(* IEC 61131-3 sources: AutoPLC/data/rag_data/st/st_case_code (part 2) *)

(* ---- ELEMENT_GET.st ---- *)
FUNCTION ELEMENT_GET : string
VAR_INPUT
    SEP : BYTE;
    POS : INT;
END_VAR

VAR_IN_OUT
    ELEMENT : STRING[ELEMENT_LENGTH];
END_VAR_IN_OUT

VAR
    i : INT := 1;
    o : INT := 1;
    pt : POINTER TO ARRAY[1..ELEMENT_LENGTH] OF BYTE;
    po : POINTER TO ARRAY[1..ELEMENT_LENGTH] OF BYTE;
    cnt : INT;
    c : BYTE;
END_VAR
(* load pointers *)
pt := ADR(ELEMENT);
po := ADR(ELEMENT_GET);

(* search for the n-th occurence of a separation character and store position in i *)
WHILE (cnt < pos) AND (i < ELEMENT_LENGTH) AND (pt^[i] > 0) DO
	IF pt^[i] = sep THEN cnt := cnt + 1; END_IF;
	i := i + 1;
END_WHILE;

(* copy the list element to output *)
IF i < ELEMENT_LENGTH THEN c := pt^[i]; END_IF;
WHILE (c <> sep) AND (c > 0) AND (o < ELEMENT_LENGTH) AND (i < ELEMENT_LENGTH) DO
	po^[o] :=pt^[i];
	o := o + 1;
	i := i + 1;
	c := pt^[i];
END_WHILE;

(* terminate the output string *)
po^[o] := 0;

(* revision histroy
ks 05. apr. 2011	rev 1.0
	original release

*)
END_FUNCTION

(* ---- ELLIPSE_A.st ---- *)
FUNCTION ELLIPSE_A : REAL
VAR_INPUT
    R1: REAL;
    R2: REAL;
END_VAR
ELLIPSE_A := math.PI * R1 * R2;

(* revision histroy
hm	16. oct 2007	rev 1.0
	original version

hm	18. oct. 2008	rev 1.1
	using math constants
*)
END_FUNCTION

(* ---- ELLIPSE_C.st ---- *)
FUNCTION ELLIPSE_C : REAL
VAR_INPUT
    R1 : REAL;
    R2 : REAL;
END_VAR
ELLIPSE_C := math.PI * (3.0 * (R1+R2) - SQRT((3.0 * r1 + R2) * (3.0 * r2 + r1)));

(* revision histroy
hm	16. oct 2007	rev 1.0
	original version

hm	18. oct. 2008	rev 1.1
	using math constants

hm	10. mar. 2009	rev 1.2
	changed syntax of real constants to 0.0

*)
END_FUNCTION

(* ---- ERF.st ---- *)
FUNCTION ERF : REAL
VAR_INPUT
    X : REAL;
END_VAR_INPUT

VAR
    x2 : REAL;
    ax2 : REAL;
END_VAR
x2 := X*X;
ax2 := 0.147 * x2 + 1.0;
ERF := SQRT(1.0 - EXP(-X2 * ((0.27323954473516 + aX2)/(ax2)))) * SGN(x);

(* revision history
hm	7. apr. 2008	rev 1.0
	original version

hm	30. jun. 2008	rev 1.1
	added type conversions to avoid warnings under codesys 3.0

hm	25. oct. 2008	rev 1.2
	new code using new algorithm

hm	10. mar. 2009	rev 1.3
	real constants updated to new systax using dot
*)
END_FUNCTION

(* ---- ERFC.st ---- *)
FUNCTION ERFC : REAL
VAR_INPUT
    X : REAL;
END_VAR
ERFC := 1.0 - ERF(X);

(* revision history
hm	7. apr. 2008	rev 1.0
	original version

hm	10. mar. 2009	rev 1.1
	real constants updated to new systax using dot

*)
END_FUNCTION

(* ---- EVEN.st ---- *)
FUNCTION EVEN : BOOL
VAR_INPUT
    in : DINT; // Input variable declaration
END_VAR
EVEN := NOT in.0;

(* revision history
hm	1. oct 2006	rev 1.0
	ORIGINAL VERSION

hm	01.12.2007	rev 1.1
	changed code for improved performance

hm	21. mar. 2008	rev 1.2
	changed type of input IN from INT to DINT
*)
END_FUNCTION

(* ---- EXEC.st ---- *)
FUNCTION EXEC : string
VAR_INPUT
    str : STRING[STRING_LENGTH];
END_VAR

VAR
    pos : INT;
    R1 : REAL;
    R2 : REAL;
    operator : STRING[10];
END_VAR
(* extract both numbers and operator *)
EXEC := UPPERCASE(TRIM(str));

pos := FINDB_NONUM(EXEC);
IF pos > 1 THEN R1 := STRING_TO_REAL(LEFT(EXEC,pos-1)); END_IF;
R2 := STRING_TO_REAL(RIGHT(EXEC,LEN(EXEC)-pos));
EXEC := LEFT(EXEC,pos);
pos := FINDB_NUM(EXEC);
operator := RIGHT(EXEC,LEN(EXEC) - pos);
IF operator = '' AND LEN(str) = 0 THEN
	EXEC := '';
	RETURN;
ELSIF operator = '' THEN
	EXEC := str;
	RETURN;
END_IF;
IF operator = '^' THEN
	EXEC := REAL_TO_STRING(EXPT(R1, R2));
ELSIF operator = 'SQRT' THEN
	EXEC := REAL_TO_STRING(SQRT(R2));
ELSIF operator = 'SIN' THEN
	EXEC := REAL_TO_STRING(SIN(r2));
ELSIF operator = 'COS' THEN
	EXEC := REAL_TO_STRING(COS(r2));
ELSIF operator = 'TAN' THEN
	EXEC := REAL_TO_STRING(TAN(R2));
ELSIF operator = '*' THEN
	EXEC := REAL_TO_STRING(R1 * R2);
ELSIF operator = '/' THEN
	IF R2 <> 0 THEN EXEC := REAL_TO_STRING(R1 / R2); ELSE EXEC := 'ERROR'; END_IF;
ELSIF operator = '+' THEN
	EXEC := REAL_TO_STRING(r1 + r2);
ELSIF operator = '-' THEN
	EXEC := REAL_TO_STRING(r1 - r2);
ELSE
	EXEC := 'ERROR';
END_IF;

IF EXEC = 'ERROR' THEN
	RETURN;
(* some systems deliver integer instead of real *)
ELSIF FIND(EXEC,'.') = 0 THEN
	EXEC := CONCAT(EXEC, '.0');
(* some systems deliver n. instead of n.0 ! *)
ELSIF RIGHT(EXEC,1) = '.' THEN
	EXEC := CONCAT(EXEC,'0');
END_IF;

(* revision history

hm 	6.feb 2007		rev 1.1
	cos has to be written in uppercase
	divide by 0 will return an error

hm	5. mar. 2008	rev 1.2
	add a 0 to the string if a '.' is at the end of the string

hm	20. mar. 2008	rev 1.3
	make sure the function always returns a real value in the form of x.y

hm	29. mar. 2008	rev 1.4
	changed STRING to STRING(STRING_LENGTH)
*)
END_FUNCTION

(* ---- EXP10.st ---- *)
FUNCTION EXP10 : REAL
VAR_INPUT
    X : REAL;
END_VAR
EXP10 := EXP(X * 2.30258509299405);

(* revision history
hm	2. dec 2007		rev 1.0
	original version

*)
END_FUNCTION

(* ---- EXPN.st ---- *)
FUNCTION EXPN : REAL
VAR_INPUT
    X : REAL;  // Input variable of type REAL
    N : INT;   // Input variable of type INT
END_VAR

VAR
    sign : BOOL;  // Local variable of type BOOL
END_VAR
sign := n.15;
N := ABS(N);
IF N.0 THEN EXPN := X; ELSE EXPN := 1.0; END_IF;
N := SHR(N,1);
WHILE N > 0 DO
   X := X * X;
   IF N.0 THEN EXPN := EXPN * X; END_IF;
   N := SHR(N,1);
END_WHILE;
IF sign THEN EXPN := 1.0 / EXPN; END_IF;

(* revision history
hm	4. dec 2007	rev 1.0
	original version

hm	22. oct. 2008	rev 1.1
	optimized code

hm	10. mar. 2009	rev 1.2
	removed nested comments
	real constants updated to new systax using dot

*)
END_FUNCTION

(* ---- F_LIN.st ---- *)
FUNCTION F_LIN : REAL
VAR_INPUT
    X : REAL;
    A : REAL;
    B : REAL;
END_VAR
F_lin := A * X + B;
END_FUNCTION

(* ---- F_LIN2.st ---- *)
FUNCTION F_LIN2 : REAL
VAR_INPUT
    X   : REAL;
    X1  : REAL;
    Y1  : REAL;
    X2  : REAL;
    Y2  : REAL;
END_VAR
F_LIN2 := (Y2 - Y1) / (X2 - X1) * (X - X1) + Y1;

(* revision history
hm	1. jan. 2007	rev 1.0
	original release

hm	17. dec. 2008	rev 1.1
	optimized formula

*)
END_FUNCTION

(* ---- F_POLY.st ---- *)
FUNCTION F_POLY : REAL
VAR_INPUT
    X : REAL;
    C : ARRAY[0..7] OF REAL;
END_VAR
F_POLY := ((((((( c[7] * x + c[6] ) * x + c[5] ) * x + c[4] ) * x + c[3] ) * x + c[2] ) * x + c[1] ) * x + c[0] ) ;

(* revision history
hm		20. may. 2008		rev 1.0
	original version

hm	18. mar. 2011	rev 1.1
	improved performance
*)
END_FUNCTION

(* ---- F_POWER.st ---- *)
FUNCTION F_POWER : REAL
VAR_INPUT
    a : REAL;
    x : REAL;
    n : REAL;
END_VAR
F_POWER := a * EXPT(X, N);
END_FUNCTION

(* ---- F_QUAD.st ---- *)
FUNCTION F_QUAD : REAL
VAR_INPUT
    X : REAL;
    A : REAL;
    B : REAL;
    C : REAL;
END_VAR
F_QUAD :=  (A * X + B) * X + C;

(* revision history

hm	1. sep. 2006	rev 1.0
	original version

hm	18. mar. 2001	rev 1.1
	improved performance
*)
END_FUNCTION

(* ---- F_TO_C.st ---- *)
FUNCTION F_TO_C : REAL
VAR_INPUT
    fahrenheit : REAL;
END_VAR
F_TO_C := (fahrenheit - 32.0) * 0.5555555555555;

(* revision history
hm	4. aug 2006	rev 1.0
	original version

hm	11. mar. 2009	rev 1.1
	real constants updated to new systax using dot

*)
END_FUNCTION

(* ---- F_TO_OM.st ---- *)
FUNCTION F_TO_OM : REAL
VAR_INPUT
    F : REAL;
END_VAR
F_TO_OM := math.PI2 * F;

(* revision history
hm	22. jan. 2007	rev 1.0
	original version

hm	18. oct. 2008	rev 1.1
	unsing math constants

*)
END_FUNCTION

(* ---- F_TO_PT.st ---- *)
FUNCTION F_TO_PT : TIME
VAR_INPUT
    F : REAL;
END_VAR
F_TO_PT := DWORD_TO_TIME(REAL_TO_DWORD(1.0 / F * 1000.0));

(* revision history

hm	4. aug. 2006	rev 1.0
	original version

hm	11. mar. 2009	rev 1.1
	real constants updated to new systax using dot

*)
END_FUNCTION

(* ---- FACT.st ---- *)
FUNCTION FACT : DINT
VAR_INPUT
    X : INT;
END_VAR
IF X >= 0 AND X <= 12 THEN
	FACT := math.FACTS[X];
ELSE
	FACT := -1;
END_IF;

(* working code without array
IF X > 12 OR X < 0 THEN
	FACT := -1;
ELSIF X < 7 THEN
	FACT := 1;
	FOR i := 2 TO X DO
		FACT := FACT * i;
	END_FOR;
ELSE
	FACT := 5040;
	FOR i := 8 TO X DO
		FACT := FACT * i;
	END_FOR;
END_IF;
*)

(* revision history
hm 4.3.2007		rev 1.1
	changed a critical error where while loop was indefinite.

hm	10.12.2007	rev 1.2
	start value for i has changed to 2 for better performance

hm	10. mar 2008	rev 1.3
	changed output of fact to dint to allow bigger values

hm	27. oct. 2008	rev 1.4
	optimized code

hm	26. mar. 2011	rev 1.5
	using array math.facts
*)
END_FUNCTION

(* ---- FIB.st ---- *)
FUNCTION FIB : DINT
VAR_INPUT
    X : INT;
END_VAR

VAR
    t1 : DINT;
    t2 : DINT;
END_VAR
IF X < 0 OR X > 46 THEN
	FIB := -1;
ELSIF x < 2 THEN
	FIB := X;
	RETURN;
ELSE
	(* the fibonacci number is the sum of the two suceeding fibonaci numbers *)
	(* we store the numbers alternatively in t1 and t2 depending on pt *)
	t2 := 1;
	WHILE X > 3 DO
		X := X-2;
		t1 := t1 + t2;
		t2 := t1 + t2;
	END_WHILE;
	IF X > 2 THEN t1 := t1 + t2; END_IF;
	fib := t1 + t2;
END_IF;

(* alternative code for very big numbers

IF X < 31 THEN
	fib := 0.4472136 * (expn(1.618034,X) - expn(-0.618034,X));
ELSE
	fib := 0.4472133 * expn(1.618034,X);
END_IF;

*)

(* revision history
hm		27. dec 2007	rev 1.0
	original version

hm		2. jan 2008	rev 1.1
	deleted unused variable pt

hm		10. mar 2008	rev 1.2
	changed output to dint instead of real

hm		26. mar. 2008	rev 1.3
	function now returns -1 for input < 0 or > 46

*)
END_FUNCTION

(* ---- FILE_BLOCK_DEMO.st ---- *)
FUNCTION FILE_BLOCK_DEMO
VAR
    PT : NETWORK_BUFFER;
    fsd : FILE_SERVER_DATA;
    FILE_SERVER : FILE_SERVER;
    FILE_BLOCK : FILE_BLOCK;
    filename : STRING := 'config.ini';
    data : BYTE;
    error : BYTE;
    mode : BYTE;
    pos : UDINT;
END_VAR

END_FUNCTION

(* ---- FILE_PATH_SPLIT.st ---- *)
FUNCTION FILE_PATH_SPLIT : BOOL
VAR_INPUT
    FILENAME : STRING[OSCAT_BASIC.STRING_LENGTH];
END_VAR

VAR_IN_OUT
    X : FILE_PATH_DATA;
END_VAR

VAR
    b : INT;
    c : INT;
    d : STRING[1];
    p1 : INT;
    p2 : INT;
END_VAR
X.DRIVE := '';
X.DIRECTORY := '';
X.FILENAME := '';
c := LEN(FILENAME);
IF c = 0 THEN
	FILE_PATH_SPLIT := FALSE;
	RETURN;
END_IF;

FOR b := 1 TO c DO
	d := MID(FILENAME, 1, b);
	IF d = ':' THEN
		p1 := b;
	ELSIF d = '/' OR d = '\' THEN
		p2 := b;
	END_IF;
END_FOR;

IF p1 = 2 THEN
	X.DRIVE := LEFT(FILENAME,p1);
END_IF;

IF p2 > 0 AND p2 > p1 THEN
	X.DIRECTORY := MID(FILENAME,p2 - p1,p1+1); (* len , pos *)
END_IF;

X.FILENAME := RIGHT(FILENAME,c - MAX (p1,p2));
FILE_PATH_SPLIT := TRUE;

(* revision history
ks	01. jan. 2011	rev 1.0
	original version
*)
END_FUNCTION

(* ---- FILL.st ---- *)
FUNCTION FILL : string
VAR_INPUT
    C : BYTE;
    L : INT;
END_VAR

VAR
    i : INT;
    sx : STRING[1];
END_VAR
Sx := CHR_TO_STRING(c);
(* limit L to maximum 80 characters the length of a standard string *)
L := LIMIT(0,L,STRING_LENGTH);
(* create a string of characters to be connected to str *)
FOR i := 1 TO 8 DO
	FILL := CONCAT(FILL,FILL);
	IF L.7 THEN FILL := CONCAT(FILL,Sx); END_IF;
	L := SHL(L,1);
END_FOR;

(* revision histroy
hm	29. mar. 2008	rev 1.0
	original release

hm	17. dec. 2008	rev 1.1
	changed function chr to chr_to_string

*)
END_FUNCTION

(* ---- FIND_CHAR.st ---- *)
FUNCTION FIND_CHAR : INT
VAR_INPUT
    str : STRING(STRING_LENGTH);
    pos : INT;
END_VAR

VAR
    i : INT;
    pt : POINTER TO ARRAY [1..255] OF BYTE;
    stop : INT;
    X : BYTE;
END_VAR
pt := ADR(str);
stop := LEN(str);
FOR i := MAX(pos,1) TO stop DO;
	X := pt^[i];
	IF X > 31 AND ((setup.EXTENDED_ASCII AND X <> 127) OR (NOT setup.EXTENDED_ASCII AND X < 127)) THEN
		FIND_CHAR := i;
		RETURN;
	END_IF;
END_FOR;
FIND_CHAR := 0;

(* revision history
hm	29. feb 2008	rev 1.0
	original version

hm	26. mar. 2008	rev 1.1
	char will now accept extended ascii

hm	29. mar. 2008	rev 1.2
	changed STRING to STRING(STRING_LENGTH)

hm	21. oct. 2008	rev 1.3
	changes setup constants
	optimized code
*)
END_FUNCTION

(* ---- FIND_CTRL.st ---- *)
FUNCTION FIND_CTRL : INT
VAR_INPUT
    str : STRING(STRING_LENGTH);
    pos : INT;
END_VAR

VAR
    i : INT;
    pt : POINTER TO ARRAY[1..255] OF BYTE;
    stop : INT;
    x : BYTE;
END_VAR
pt := ADR(str);
stop := LEN(str);
FOR i := MAX(pos,1) TO stop DO;
	x := PT^[I];
	IF x < 32 OR X = 127 THEN
		FIND_CTRL := i;
		RETURN;
	END_IF;
END_FOR;
FIND_CTRL := 0;

(* revision history
hm	29. feb 2008	rev 1.0
	original version

hm	26. mar. 2008	rev 1.1
	character 127 is now recognized as control

hm	29. mar. 2008	rev 1.2
	changed STRING to STRING(STRING_LENGTH)
*)
END_FUNCTION

(* ---- FIND_NONUM.st ---- *)
FUNCTION FIND_NONUM : INT
VAR_INPUT
    str : STRING(STRING_LENGTH);
    pos : INT;
END_VAR

VAR
    i : INT;
    pt : POINTER TO ARRAY[1..255] OF BYTE;
    end : INT;
    X : BYTE;
END_VAR
pt := ADR(str);
end := LEN(str);
FOR i := MAX(pos,1) TO end DO;
	X := pt^[i];
	IF (X < 48 AND X <> 46) OR X > 57 THEN
		FIND_NONUM := i;
		RETURN;
	END_IF;
END_FOR;
FIND_NONUM := 0;

(* revision history
hm	6. oct. 2006	rev 1.0
	original version

hm	29. feb 2008	rev 1.1
	added input pos to start search at position

hm	29. mar. 2008	rev 1.2
	changed STRING to STRING(STRING_LENGTH)

hm	21. oct. 2008	rev 1.3
	optimized code

*)
END_FUNCTION

(* ---- FIND_NUM.st ---- *)
FUNCTION FIND_NUM : INT
VAR_INPUT
    str : STRING(SIZE := STRING_LENGTH);
    pos : INT;
END_VAR

VAR
    i : INT;
    pt : POINTER TO ARRAY[1..255] OF BYTE;
    stop : INT;
    X : BYTE;
END_VAR
pt := ADR(str);
stop := LEN(str);
FOR i := MAX(pos,1) TO stop DO;
	X := pt^[i];
	IF (X > 47 AND X < 58) OR X = 46 THEN
		FIND_NUM := i;
		RETURN;
	END_IF;
END_FOR;
FIND_NUM := 0;

(* revision history
hm	6. oct. 2006	rev 1.0
	original version

hm	29. feb 2008	rev 1.1
	added input pos to start search at position

hm	29. mar. 2008	rev 1.2
	changed STRING to STRING(STRING_LENGTH)

*)
END_FUNCTION

(* ---- FINDB.st ---- *)
FUNCTION FINDB : INT
VAR_INPUT
    str1 : STRING(STRING_LENGTH);
    str2 : STRING(STRING_LENGTH);
END_VAR

VAR
    pos : INT;
    length : INT;
END_VAR
length := LEN(str2);
FOR pos := LEN(str1) - length + 1 TO 1 BY -1 DO
	IF MID(str1,length,pos) = str2 THEN
		FindB := pos;
		RETURN;
	END_IF;
END_FOR;
FindB := 0;

(* revision history
hm	6. oct 2006		rev 1.0
	original version

hm	15 dec 2007		rev 1.1
	changed code for better performance

hm	29. feb 2008	rev 1.2
	added findb := 0 for compatibility reasons

hm	29. mar. 2008	rev 1.3
	changed STRING to STRING(STRING_LENGTH)
*)
END_FUNCTION

(* ---- FINDB_NONUM.st ---- *)
FUNCTION FINDB_NONUM : INT
VAR_INPUT
    str : STRING(STRING_LENGTH);
END_VAR

VAR
    pos : INT;
    pt : POINTER TO BYTE;
END_VAR
pt := ADR(str) + LEN(str) - 1;
FOR pos := LEN(str) TO 1 BY -1 DO;
	IF (PT^ < 48 AND PT^ <> 46) OR PT^ > 57 THEN
		FINDB_NONUM := pos;
		RETURN;
	END_IF;
	PT := PT - 1;
END_FOR;
FINDB_NONUM := 0;

(* revision history
hm	6. oct 2006		rev 1.0
	original version

hm	29. feb 2008	rev 1.1
	improved performance

hm	29. mar. 2008	rev 1.2
	changed STRING to STRING(STRING_LENGTH)

hm	21. oct. 2008	rev 1.3
	optimized code
*)
END_FUNCTION

(* ---- FINDB_NUM.st ---- *)
FUNCTION FINDB_NUM : INT
VAR_INPUT
    str : STRING:= STRING_LENGTH; // Input variable of type STRING with specified length
END_VAR

VAR
    pos : INT; // Local variable of type INT
    pt : POINTER TO BYTE; // Local variable of type pointer to BYTE
END_VAR
pt := ADR(str) + LEN(str) - 1;
FOR pos := LEN(str) TO 1 BY -1 DO;
	IF (PT^ > 47 AND PT^ < 58) OR PT^ = 46 THEN
		FINDB_NUM := pos;
		RETURN;
	END_IF;
	PT := PT - 1;
END_FOR;
FINDB_NUM := 0;

(* revision history
hm	6. oct 2006		rev 1.0
	original version

hm	29. feb 2008	rev 1.1
	improved performance

hm	29. mar. 2008	rev 1.2
	changed STRING to STRING(STRING_LENGTH)
*)
END_FUNCTION

(* ---- FINDP.st ---- *)
FUNCTION FINDP : INT
VAR_INPUT
    str : STRING[STRING_LENGTH];
    src : STRING[STRING_LENGTH];
    pos : INT;
END_VAR

VAR
    i : INT;
    ls : INT;
    lx : INT;
    stp : INT;
END_VAR
ls := LEN(str);
lx := LEN(src);
IF ls < lx OR lx = 0 THEN RETURN; END_IF;
stp := ls - lx + 1;
FOR i := MAX(pos,1) TO stp DO
	IF MID(str,lx,i) = src THEN
		FINDP := i;
		RETURN;
	END_IF;
END_FOR;
FINDP := 0;

(* revision histroy
hm	4. feb. 2008	rev 1.0
	original release

hm	29. feb 2008	rev 1.1
	ADDED MAX(pos,1) in loop initialization

hm	29. mar. 2008	rev 1.2
	changed STRING to STRING(STRING_LENGTH)
*)
END_FUNCTION

(* ---- FIX.st ---- *)
FUNCTION FIX : string
VAR_INPUT
    str : STRING[STRING_LENGTH];
    L : INT;
    C : BYTE;
    M : INT;
END_VAR

VAR
    N : INT;
    SX : STRING[STRING_LENGTH];
END_VAR
(* make sure L does not exceed the limits of a string *)
N := LIMIT(0,L,STRING_LENGTH) - LEN(str);
IF N <= 0 THEN
	(* truncate the string at length N *)
	IF M = 1 THEN
		FIX := RIGHT(str,L);
	ELSE
		FIX := LEFT(str,L);
	END_IF;
ELSIF M = 1 THEN
	(* connect fill characters at the beginning *)
	sx := FILL(C,N);
	FIX := CONCAT(sx,str);
ELSIF M = 2 THEN
	(* center str beween fill characters *)
	(* for an uneven number of fill characters, there is one more at the end *)
	sx := FILL(C,SHR(N+1,1));
	FIX := CONCAT(str,sx);
	SX := LEFT(sx,SHR(N,1));
	FIX := CONCAT(sx,FIX);
ELSE
	(* connect fill characters at the end *)
	SX := FILL(C,N);
	FIX := CONCAT(str,SX);
END_IF;

(* revision histroy
hm	29. mar. 2008	rev 1.0
	original release

*)
END_FUNCTION

(* ---- FLOAT_TO_REAL.st ---- *)
FUNCTION FLOAT_TO_REAL : REAL
VAR_INPUT
    FLT : STRING[20];
END_VAR

VAR
    pt : POINTER TO ARRAY[1..20] OF BYTE;
    i : INT;
    X : BYTE;
    sign : INT := 1;
    stop : INT;
    tmp : DINT;
    d : INT;
END_VAR
pt := ADR(FLT);
stop := LEN(FLT);

(* we first check for sign and exit if first number or dot is reached *)
FOR i := 1 TO stop DO
	X := pt^[i];
	IF X > 47 AND X < 58 OR X = 46 THEN
		EXIT;
	ELSIF X = 45 THEN
		(* code 45 is sign *)
		sign := -1;
	END_IF;
END_FOR;

(* now we scan numbers till end or dot or E is reached *)
FOR i := i TO stop DO
	X := pt^[i];
	IF X = 44 OR X = 46 OR X = 69 OR X = 101 THEN
		EXIT;
	(* calculate the value of the digit *)
	ELSIF X > 47 AND x < 58 THEN
		tmp := tmp * 10 + X - 48;
	END_IF;
END_FOR;

(* process the portion after the comma if comma or dot is reached exit if exponent starts *)
IF x = 44 OR X = 46 THEN
	FOR i := i + 1 TO stop DO
		X := pt^[i];
		IF X = 69 OR X = 101 THEN
			EXIT;
		ELSIF x > 47 AND x < 58 THEN
			tmp := tmp * 10 + X - 48;
			d := d - 1;
		END_IF;
	END_FOR;
END_IF;

(* process exponent if present *)
IF X = 69 OR X = 101 THEN
	d := d + DEC_TO_INT(RIGHT(FLT, stop - i));
END_IF;

FLOAT_TO_REAL :=  EXPN(10, d) * DINT_TO_REAL(TMP * SIGN);

(* revision histroy
hm	22. jun. 2008	rev 1.0
	original release

hm	2. oct. 2008	rev 1.1
	fixed an error, characters 8 and 9 would not be converted

hm	22. oct. 2008	rev 1.2
	last fix was not done correctly

hm	23. oct. 2008	rev 1.3
	optimzed code
*)
END_FUNCTION

(* ---- FLOOR.st ---- *)
FUNCTION FLOOR : INT
VAR_INPUT
    X : REAL;
END_VAR
FLOOR := REAL_TO_INT(X);
IF FLOOR > X THEN
	FLOOR := FLOOR - 1;
END_IF;

(* revision history
hm		7. feb 2007		rev 1.0
	originlal version

hm		21. mar. 2008	rev 1.1
	replaced trunc with real_to_int for compatibility reasons

*)
END_FUNCTION

(* ---- FLOOR2.st ---- *)
FUNCTION FLOOR2 : DINT
VAR_INPUT
    X : REAL;
END_VAR
FLOOR2 := REAL_TO_DINT(X);
IF DINT_TO_REAL(FLOOR2) > X THEN
	FLOOR2 := FLOOR2 - 1;
END_IF;

(* revision history
hm	21. mar. 2008	rev 1.0
	originlal version

hm	4. apr. 2008	rev 1.1
	added type conversion to avoid warnings under codesys 3.0
*)
END_FUNCTION

(* ---- FRACT.st ---- *)
FUNCTION FRACT : REAL
VAR_INPUT
    x : REAL;
END_VAR
IF ABS(x) < 2.0E9 THEN
	FRACT := x - DINT_TO_REAL(D_TRUNC(x));
ELSE
	FRACT := 0.0;
END_IF;

(* revision history
hm	4. aug 2006	rev 1.0
	original version

hm	11. mar 2008	rev 1.1
	added dint_to_real for compatibility reasons
	now returns 0 for number > 2e9
	changed input to x

hm	21. mar. 2008	rev 1.2
	use D_trunc instead of TRUNC for compatibility reasons

hm	10. mar. 2009	rev 1.3
	real constants updated to new systax using dot

*)
END_FUNCTION

(* ---- FRMP_B.st ---- *)
FUNCTION FRMP_B : BYTE
VAR_INPUT
    START : BYTE;
    DIR   : BOOL;
    TD    : TIME;
    TR    : TIME;
END_VAR
IF TD < TR THEN
	FRMP_B := MIN(DWORD_TO_BYTE(SHL(TIME_TO_DWORD(TD), 8) / TIME_TO_DWORD(TR)), SEL(DIR, START, BYTE#255 - START));
	IF DIR THEN
		FRMP_B := START + FRMP_B;
	ELSE
		FRMP_B := START - FRMP_B;
	END_IF;
ELSE
	FRMP_B := SEL(DIR, 0, 255);
END_IF;

(* revision history

17. feb. 2011	rev 1.0
	new module

*)
END_FUNCTION

(* ---- FSTRING_TO_BYTE.st ---- *)
FUNCTION FSTRING_TO_BYTE : BYTE
VAR_INPUT
    IN: STRING[12];
END_VAR
IF LEFT(IN, 2) = '2#' THEN
	(* we need to convert binary *)
	FSTRING_TO_BYTE := BIN_TO_BYTE(RIGHT(in, LEN(in) - 2));
ELSIF LEFT(in, 2) = '8#' THEN
	(* weneed to convert octals *)
	FSTRING_TO_BYTE := OCT_TO_BYTE(RIGHT(in, LEN(in) - 2));
ELSIF LEFT(in, 3) = '16#' THEN
	(* we need to convert hexadecimal *)
	FSTRING_TO_BYTE := HEX_TO_BYTE(RIGHT(in, LEN(in) - 3));
ELSE
	(* we assume decimal representation *)
	FSTRING_TO_BYTE := DEC_TO_BYTE(CLEAN(in,'0123456789'));
END_IF;

(* revision histroy
hm	18. jun. 2008	rev 1.0
	original release

hm	20. sep. 2008	rev 1.1
	changed length of input string from 20 to 12
*)
END_FUNCTION

(* ---- FSTRING_TO_DT.st ---- *)
FUNCTION FSTRING_TO_DT : DT
VAR_INPUT
    SDT: STRING[60];    // Input variable for source data text
    FMT: STRING[60];    // Input variable for format
END_VAR

VAR CONSTANT
    ignore: STRING[1] := '*';  // ignore character is *
    fchar: STRING[1] := '#';    // format character is #
END_VAR

VAR
    c: STRING[1];    // local variable for character
    tmp: STRING[20];  // local variable for temporary storage
    end: INT;         // local variable for end indicator
    dy: INT := 1970;  // local variable for year, initialized to 1970
    dm: INT := 1;     // local variable for month, initialized to 1
    dd: INT := 1;     // local variable for day, initialized to 1
    th: INT;         // local variable for hour
    tm: INT;         // local variable for minute
    ts: INT;         // local variable for second
END_VAR
(* scan input string *)
WHILE fmt <> '' DO
	c := LEFT(fmt,1);
	IF c = ignore THEN
		(* skip ignore characters *)
		fmt := DELETE(fmt,1,1);
		sdt := DELETE(sdt,1,1);
	ELSIF C = fchar THEN
		(* format chracter found skip format char and read identifier *)
		(* store format identifier in c and skip to next char in fmt *)
		c := MID(fmt,1,2);
		fmt := DELETE(fmt,2,1);
		(* extract the substring until the end of sdt or to next char of fmt *)
		IF fmt = '' THEN
			tmp := sdt;
		ELSE
			(* serach for end of substring *)
			end := FIND(sdt, LEFT(fmt,1))-1;
			tmp := LEFT(sdt, end);
			sdt := DELETE(sdt, end,1);
		END_IF;
		(* extract information from substring *)
		IF c = 'Y' THEN
			dy := STRING_TO_INT(tmp);
			IF dy < 100 THEN dy := dy + 2000; END_IF;
		ELSIF c = 'M' THEN
			dm := STRING_TO_INT(tmp);
		ELSIF c = 'N' THEN
			dm := FSTRING_TO_MONTH(tmp,0);
		ELSIF c = 'D' THEN
			dd := STRING_TO_INT(tmp);
		ELSIF c = 'h' THEN
			th := STRING_TO_INT(tmp);
		ELSIF c = 'm' THEN
			tm := STRING_TO_INT(tmp);
		ELSIF c = 's' THEN
			ts := STRING_TO_INT(tmp);
		END_IF;
	ELSIF c = LEFT(sdt,1) THEN
		(* skip matching characters *)
		fmt := DELETE(fmt,1,1);
		sdt := DELETE(sdt,1,1);
	ELSE
		RETURN;
	END_IF;
END_WHILE;

FSTRING_TO_DT := SET_DT(dy,dm,dd,th,tm,ts);

(* revision histroy
hm	24. sep. 2008	rev 1.0
	original release

*)
END_FUNCTION

(* ---- FSTRING_TO_DWORD.st ---- *)
FUNCTION FSTRING_TO_DWORD : DWORD
VAR_INPUT
    IN : STRING[40];
END_VAR
IF LEFT(IN, 2) = '2#' THEN
	(* we need to convert binary *)
	FSTRING_TO_DWORD := BIN_TO_DWORD(RIGHT(in, LEN(in) - 2));
ELSIF LEFT(in, 2) = '8#' THEN
	(* weneed to convert octals *)
	FSTRING_TO_DWORD := OCT_TO_DWORD(RIGHT(in, LEN(in) - 2));
ELSIF LEFT(in, 3) = '16#' THEN
	(* we need to convert hexadecimal *)
	FSTRING_TO_DWORD := HEX_TO_DWORD(RIGHT(in, LEN(in) - 3));
ELSE
	(* we assume decimal representation *)
	FSTRING_TO_DWORD := DEC_TO_DWORD(CLEAN(in,'0123456789'));
END_IF;

(* revision histroy
hm	18. jun. 2008	rev 1.0
	original release

hm	20. sep. 2008	rev 1.1
	changed length of input dtring from 20 to 40

*)
END_FUNCTION

(* ---- FSTRING_TO_MONTH.st ---- *)
FUNCTION FSTRING_TO_MONTH : INT
VAR_INPUT
    MTH : STRING(20);
    LANG : INT;
END_VAR

VAR
    lx : INT;
END_VAR
IF LANG = 0 THEN lx := LANGUAGE.DEFAULT; ELSE lx := MIN(LANG, LANGUAGE.LMAX); END_IF;
MTH := TRIM(mth);
MTH := CAPITALIZE(LOWERCASE(MTH));

FOR FSTRING_TO_MONTH := 1 TO 12 DO
	IF MTH = language.MONTHS[lx, FSTRING_TO_MONTH] THEN RETURN; END_IF;
	IF MTH = language.MONTHS3[lx, FSTRING_TO_MONTH] THEN RETURN; END_IF;
END_FOR;

(* since no name matched try to decode as integer *)
FSTRING_TO_MONTH := STRING_TO_INT(MTH);

(* revision histroy
hm	25. sep. 2008	rev 1.0
	original release

hm	19. oct. 2008	rev 1.1
	changed language setup constants

hm	25. oct. 2008	rev 1.2
	optimized code
*)
END_FUNCTION

(* ---- FSTRING_TO_WEEK.st ---- *)
FUNCTION FSTRING_TO_WEEK : BYTE
VAR_INPUT
    WEEK : STRING[60];
    LANG : INT;
END_VAR

VAR
    pos : INT;
END_VAR
pos := FIND(WEEK, ',');
WHILE pos > 0 DO
	FSTRING_TO_WEEK := FSTRING_TO_WEEK OR SHR(BYTE#128, FSTRING_TO_WEEKDAY(MID(WEEK, pos - 1, 1), LANG));
	WEEK := RIGHT(WEEK, LEN(Week) - pos);
	pos := FIND(WEEK, ',');
END_WHILE;
FSTRING_TO_WEEK := (FSTRING_TO_WEEK OR SHR(BYTE#128, FSTRING_TO_WEEKDAY(WEEK, LANG))) AND BYTE#127;

(* revision histroy
hm	18. jun. 2008	rev 1.0
	original release

hm	25. oct. 2008	rev 1.1
	using language defauls and input lang
*)
END_FUNCTION

(* ---- FSTRING_TO_WEEKDAY.st ---- *)
FUNCTION FSTRING_TO_WEEKDAY : INT
VAR_INPUT
    WDAY : STRING[20];
    LANG : INT;
END_VAR

VAR
    tmp : STRING[2];
    i : INT;
    ly : INT;
END_VAR
IF LANG = 0 THEN ly := LANGUAGE.DEFAULT; ELSE ly := MIN(LANG, LANGUAGE.LMAX); END_IF;
(* tmp needs to be calculated first otherwise find can return wrong values *)
tmp := TRIM(wday);
tmp := CAPITALIZE(LOWERCASE(tmp));
FOR i := 1 TO 7 DO
	IF language.WEEKDAYS2[ly, i] = tmp THEN
		FSTRING_TO_WEEKDAY := i;
		RETURN;
	END_IF;
END_FOR;
FSTRING_TO_WEEKDAY := STRING_TO_INT(WDAY);

(* revision histroy
hm	18. jun. 2008	rev 1.0
	original release

hm	18. jul. 2008	rev 1.1
	changed nested call of left(trim()) for compatibility reasons

hm	25. oct. 2008	rev 1.2
	using language constants
*)
END_FUNCTION

(* ---- FTP_CLIENT_DEMO.st ---- *)
FUNCTION FTP_CLIENT_DEMO
VAR
    FTP_CLIENT : FTP_CLIENT;
    ftp_activate : BOOL;
    ftp_done : BOOL;
    ftp_busy : BOOL;
    ftp_error_c : DWORD;
    ftp_error_t : BYTE;
    ftp_url : STRING := 'ftp://581920:123456@oscat.atwebpages.com:2000/subordner/';
    ftp_filename : STRING := '0100kb.bin';
    ftp_download : BOOL := TRUE;
    ftp_activ : BOOL := FALSE;
    file_delete : BOOL := FALSE;
    ftp_timeout : TIME := TIME#30s0ms;
    zeit : TIME := TIME#30s0ms;
    stop : BOOL;
    start : BOOL := TRUE;
    reset : BOOL;
    error : DWORD;
    ok : DWORD;
    CLK_PRG_1 : oscatie_basic.CLK_PRG;
    COUNT_DR_1 : oscatie_basic.COUNT_DR;
    COUNT_DR_2 : oscatie_basic.COUNT_DR;
END_VAR

END_FUNCTION

(* ---- GAMMA.st ---- *)
FUNCTION GAMMA : REAL
VAR_INPUT
    X : REAL;
END_VAR
IF x > 0.0 THEN
	GAMMA := SQRT(math.PI2 / X) * EXPT(math.E_INV * (x + 1.0 / (12.0 * x - 0.1 / X)), X);
END_IF;

(* the stirling formula is not very accurate for small values of X
IF X >=0 THEN GAMMA := SQRT(math.PI2 * X) * EXPT(X / math.E, X); END_IF;
*)

(* revision history
hm	10.12.2007	rev 1.0
	original version

hm	18. oct. 2008	rev 1.1
	using math constants

hm	26. oct. 2008	rev 1.2
	using new formula with better accuracy

hm	10. mar. 2009	rev 1.3
	real constants updated to new systax using dot

*)
END_FUNCTION

(* ---- GAUSS.st ---- *)
FUNCTION GAUSS : REAL
VAR_INPUT
    X : REAL;
    U : REAL;
    SI : REAL;
END_VAR

VAR
    temp : REAL;
    si_inv : REAL;
END_VAR
temp := X - U;
si_inv := 1.0  / si;
GAUSS := EXP(Temp * Temp * si_inv * si_inv * - 0.5) * 0.39894228 * si_inv;

(* revision hisdtory
hm	6. apr. 2008	rev 1.0
	original version

hm	27. oct. 2008	rev 1.1
	optimized performance

hm	10. mar. 2009	rev 1.2
	real constants updated to new systax using dot

*)
END_FUNCTION

(* ---- GAUSSCD.st ---- *)
FUNCTION GAUSSCD : REAL
VAR_INPUT
    X : REAL;
    U : REAL;
    SI : REAL;
END_VAR
GAUSSCD := (ERF((X - U) / (SI * 1.414213562)) + 1.0) * 0.5;

(* revision hisdtory
hm	6. apr. 2008	rev 1.0
	original version

hm	10. mar. 2009	rev 1.1
	real constants updated to new systax using dot

*)
END_FUNCTION

(* ---- GCD.st ---- *)
FUNCTION GCD : INT
VAR_INPUT
    A : DINT;
    B : DINT;
END_VAR

VAR
    t : DINT;
END_VAR
IF A = 0 THEN
	GCD := DINT_TO_INT(ABS(B));
ELSIF B = 0 THEN
	GCD := DINT_TO_INT(ABS(A));
ELSE
	A := ABS(A);
	B := ABS(B);
	GCD := 1;
	WHILE NOT(A.0 OR B.0) DO
		A := SHR(A,1);
		B := SHR(B,1);
		GCD := SHL(GCD,1);
	END_WHILE;
	WHILE A > 0 DO
		IF NOT(A.0) THEN A := SHR(A,1);
		ELSIF NOT(B.0) THEN B := SHR(B,1);
		ELSE
			t:= SHR(ABS(A-B),1);
			IF A < B THEN B := t; ELSE A := T; END_IF;
		END_IF;
	END_WHILE;
	GCD := GCD * DINT_TO_INT(B);
END_IF;

(* revision history
hm	19. jan. 2011	rev 1.0
	original version

*)
END_FUNCTION

(* ---- GDF.st ---- *)
FUNCTION GDF : REAL
VAR_INPUT
    X : REAL;
END_VAR
IF X = 0.0 THEN
	GDF := 0.0;
ELSIF X > 15.0 THEN
	GDF := math.PI05;
ELSIF X < -15.0 THEN
	GDF := -math.PI05;
ELSE
	GDF := ATAN(EXP(X)) * 2.0 - math.PI05;
END_IF;

(* revision history
hm	27. apr. 2008	rev 1.0
	original version

hm	18. oct. 2008	rev 1.1
	using math constants

hm	10. mar. 2009	rev 1.2
	real constants updated to new systax using dot

*)
END_FUNCTION

(* ---- GEO_TO_DEG.st ---- *)
FUNCTION GEO_TO_DEG : REAL
VAR_INPUT
    D : INT;
    M : INT;
    SEC : REAL;
END_VAR
GEO_TO_DEG := INT_TO_REAL(D) + INT_TO_REAL(M) * 0.016666666666667 + sec * 0.00027777777777778;

(* revision histroy
hm	22. jan. 2009	rev 1.0
	original release

*)
END_FUNCTION

(* ---- GET_WAN_IP_DEMO.st ---- *)
FUNCTION GET_WAN_IP_DEMO
VAR
    GET_WAN_IP : GET_WAN_IP;   (* Derived type *)
    IP_C : IP_C;               (* Derived type *)
    S_BUF : NETWORK_BUFFER;     (* Derived type *)
    R_BUF : NETWORK_BUFFER;     (* Derived type *)
    IP_CONTROL_1 : IP_CONTROL;  (* Derived type *)
    activate : BOOL;           (* Boolean variable *)
    done : BOOL;               (* Boolean variable *)
    error_c : DWORD;          (* Double Word variable *)
    error_t : BYTE;           (* Byte variable *)
    wan_ip : STRING;          (* String variable *)
    new_ip : BOOL;            (* Boolean variable *)
END_VAR

END_FUNCTION

(* ---- GOLD.st ---- *)
FUNCTION GOLD : REAL
VAR_INPUT
    X : REAL;
END_VAR
GOLD := (X + SQRT(X*X + 4.0)) * 0.5;

(* revision history
hm	27. apr. 2008	rev 1.0
	original version

hm	10. mar. 2009	rev 1.1
	real constants updated to new systax using dot

*)
END_FUNCTION

(* ---- GRAY_TO_BYTE.st ---- *)
FUNCTION GRAY_TO_BYTE : BYTE
VAR_INPUT
    IN : BYTE;
END_VAR
GRAY_TO_BYTE := SHR(IN,4) XOR IN;
GRAY_TO_BYTE := SHR(GRAY_TO_BYTE,2) XOR GRAY_TO_BYTE;
GRAY_TO_BYTE := SHR(GRAY_TO_BYTE,1) XOR GRAY_TO_BYTE;

(* revision history
hm	9. nov. 2009	rev 1.0
	original version

*)
END_FUNCTION

(* ---- HEAT_INDEX.st ---- *)
FUNCTION HEAT_INDEX : REAL
VAR_INPUT
    T : REAL;
    RH : REAL;
END_VAR

VAR
    RH2 : REAL;
    T2 : REAL;
END_VAR
IF RH < 20.0 OR T < 20.0 THEN
	HEAT_INDEX := T;
ELSE
	RH2 := RH * RH;
	T := OSCAT_BASIC.C_TO_F(T);
	T2 := T * T;
	HEAT_INDEX := -42.379 + 2.04901523 * T - 6.83783E-3 * T2
			+ RH * (10.1433127 - 0.22475541 * T + 1.22874E-3 * T2)
			+ RH2 * (8.5282E-4 * T - 5.481717E-2 - 1.99E-6 * T2);
	HEAT_INDEX := OSCAT_BASIC.F_TO_C(HEAT_INDEX);
END_IF;

(* revision history

hm 27.2.2007		rev 1.1
	deleted unused variables rh3 and T3

hm	2.12.2007		rev 1.2
	changed code for better performance

hm	13. mar. 2009	rev 1.3
	real constants updated to new systax using dot

*)
END_FUNCTION

(* ---- HEX_TO_BYTE.st ---- *)
FUNCTION HEX_TO_BYTE : BYTE
VAR_INPUT
    HEX : STRING(5);
END_VAR

VAR
    pt : POINTER TO BYTE;
    i : INT;
    X : BYTE;
    stop : INT;
END_VAR
pt := ADR(hex);
stop := LEN(hex);
FOR I := 1 TO stop DO
	(* read the first character and subtract 48 to get value in decimal 0 = 48 *)
	x := pt^;
	(* calculate the value of the digit *)
	IF X > 47 AND x < 58 THEN
		HEX_TO_BYTE := SHL(HEX_TO_BYTE,4) + X - 48;
	ELSIF X > 64 AND X < 71 THEN
		HEX_TO_BYTE := SHL(HEX_TO_BYTE,4) + X - 55;
	ELSIF X > 96 AND X < 103 THEN
		HEX_TO_BYTE := SHL(HEX_TO_BYTE,4) + X - 87;
	END_IF;
	pt := pt + 1;
END_FOR;

(* revision histroy
hm	18. jun. 2008	rev 1.0
	original release

hm	20. sep.2008	rev 1.1
	changed length of input string from 20 to 5

*)
END_FUNCTION

(* ---- HEX_TO_DWORD.st ---- *)
FUNCTION HEX_TO_DWORD : DWORD
VAR_INPUT
    Hex: STRING[20];
END_VAR

VAR
    pt: POINTER TO BYTE;
    i: INT;
    X: BYTE;
    stop: INT;
END_VAR
pt := ADR(hex);
stop := LEN(hex);
FOR I := 1 TO stop DO
	(* read the first character and subtract 48 to get value in decimal 0 = 48 *)
	x := pt^;
	(* calculate the value of the digit *)
	IF X > 47 AND x < 58 THEN
		HEX_TO_DWORD := SHL(HEX_TO_DWORD,4) + X - 48;
	ELSIF X > 64 AND X < 71 THEN
		HEX_TO_DWORD := SHL(HEX_TO_DWORD,4) + X - 55;
	ELSIF X > 96 AND X < 103 THEN
		HEX_TO_DWORD := SHL(HEX_TO_DWORD,4) + X - 87;
	END_IF;
	pt := pt + 1;
END_FOR;

(* revision histroy
hm	2.10.2007		rev 1.0
	original release

hm	19.11.2007		rev 1.1
	changed type of function from int to dword

hm 	4. mar 2008		rev 1.2
	added support for a..f and return 0 for invalid string

hm	29. mar. 2008	rev 1.3
	changed STRING to STRING(8)

hm	18. jun. 2008	rev 1.4
	changed input hex to STRING(20)
	function now ignores wrong characters
*)
END_FUNCTION

(* ---- HOUR.st ---- *)
FUNCTION HOUR : INT
VAR_INPUT
    itod : TIME_OF_DAY; // Declaration of input variable itod of type TIME_OF_DAY
END_VAR
HOUR := DWORD_TO_INT(TOD_TO_DWORD(itod) / 3600000);

(* change history
hm 4. aug 2006	rev 1.0
	original version

hm 2.10.2006 	rev 1.1
	changed name of input to itod

*)
END_FUNCTION

(* ---- HOUR_OF_DT.st ---- *)
FUNCTION HOUR_OF_DT : INT
VAR_INPUT
    XDT : DT;
END_VAR
HOUR_OF_DT := DWORD_TO_INT((DT_TO_DWORD(XDT) MOD 86400) / 3600);

(* revision history
hm		6.9.2008	rev 1.0
	original version

*)
END_FUNCTION

(* ---- HOUR_TO_TIME.st ---- *)
FUNCTION HOUR_TO_TIME : TIME
VAR_INPUT
    IN : REAL;
END_VAR
HOUR_TO_TIME := DWORD_TO_TIME(REAL_TO_DWORD(IN * 3600000));

(* revision history
hm		4. aug 2006	rev 1.0
	original version

hm	14. mar. 2008	rev 1.1
	rounded the input after the last digit

hm	24. feb. 2009	rev 1.2
	changed input to IN
*)
END_FUNCTION

(* ---- HOUR_TO_TOD.st ---- *)
FUNCTION HOUR_TO_TOD : TOD
VAR_INPUT
    IN : REAL;
END_VAR
HOUR_TO_TOD := DWORD_TO_TOD(REAL_TO_DWORD(IN * 3600000));

(* revision history
hm	4. aug. 2006	rev 1.0
	original version

hm	14. mar. 2008	rev 1.1
	rounded the input after the last digit

hm	24. feb. 2009	rev 1.2
	changed input to IN
*)
END_FUNCTION

(* ---- HTML_DECODE.st ---- *)
FUNCTION HTML_DECODE : string
VAR_INPUT
    IN : STRING(OSCAT_BASIC.STRING_LENGTH);
END_VAR

VAR
    pos : INT;
    end : INT;
    tmp : STRING(10);
    code : STRING(1);
END_VAR
HTML_DECODE := IN;

(* docode characters encoded by character position *)
pos := FIND(HTML_DECODE, '&');
WHILE pos > 0 DO
	tmp := MID(HTML_DECODE, 2, pos + 1);
	IF tmp = '#x' OR tmp = '#X' THEN
		(* hexadecimal representation found *)
		tmp := MID(HTML_DECODE, 10, pos + 3);
		end := FIND(tmp, ';');
		CODE := OSCAT_BASIC.CHR_TO_STRING(DWORD_TO_BYTE(OSCAT_BASIC.HEX_TO_DWORD(LEFT(tmp, end - 1))));
		HTML_DECODE := REPLACE(HTML_DECODE, CODE, end + 3, pos);
	ELSIF LEFT(tmp,1) = '#' THEN
		tmp := MID(HTML_DECODE, 10, pos + 2);
		end := FIND(tmp, ';');
		CODE := OSCAT_BASIC.CHR_TO_STRING(INT_TO_BYTE(STRING_TO_INT(LEFT(tmp, end - 1))));
		HTML_DECODE := REPLACE(HTML_DECODE, CODE, end + 2, pos);
	ELSE
		(* replace all named characters *)
		tmp := MID(HTML_DECODE, 10, pos + 1);
		end := FIND(tmp, ';');
		CODE := OSCAT_BASIC.CHR_TO_STRING(OSCAT_BASIC.CHARCODE(LEFT(tmp, end - 1)));
		HTML_DECODE := REPLACE(HTML_DECODE, CODE, end + 1, pos);
	END_IF;
	(* search for next occurence of encoded characters *)
	pos := OSCAT_BASIC.FINDP(HTML_DECODE, '&', pos + 1);
END_WHILE;

(* revision history
hm	3. mai. 2008	rev 1.0
	original version

hm	16. jun. 2008	rev 1.1
	changed nested call of replace for better compatibility

hm	17. dec. 2008	rev 1.2
	changed function CHR to CHR_TO_STRING

hm	10. may. 2010	rev 1.3
	stringlength 250

*)
END_FUNCTION

(* ---- HTML_ENCODE.st ---- *)
FUNCTION HTML_ENCODE : string
VAR_INPUT
    IN : STRING(OSCAT_BASIC.STRING_LENGTH);
    M : BOOL;
END_VAR

VAR
    pt_in : POINTER TO ARRAY[1..255] OF BYTE;
    pt_out : POINTER TO ARRAY[1..256] OF BYTE;
    pos_in : INT;
    pos_out : INT;
    stop : INT;
    B : BYTE;
    tmp : STRING(10);
    i : INT;
END_VAR
pt_in  := ADR(in);
pt_out := ADR(HTML_ENCODE);

(* scan the input string and convert unallowed characters *)
pos_in := 1;
stop := LEN(in);
FOR pos_out := 1 TO 250 DO
	IF pos_in > stop THEN EXIT; END_IF;
	B := pt_in^[pos_in];
	CASE BYTE_TO_INT(B) OF
		34: (* " detected *)
			IF pos_out > OSCAT_BASIC.STRING_LENGTH - 6 THEN EXIT; END_IF;
			pt_out^[pos_out] := 38;
			pos_out := pos_out + 1;
			pt_out^[pos_out] := 113;
			pos_out := pos_out + 1;
			pt_out^[pos_out] := 117;
			pos_out := pos_out + 1;
			pt_out^[pos_out] := 111;
			pos_out := pos_out + 1;
			pt_out^[pos_out] := 116;
			pos_out := pos_out + 1;
			pt_out^[pos_out] := 59;
		38: (* & detected *)
			IF pos_out > OSCAT_BASIC.STRING_LENGTH - 5 THEN EXIT; END_IF;
			pt_out^[pos_out] := 38;
			pos_out := pos_out + 1;
			pt_out^[pos_out] := 97;
			pos_out := pos_out + 1;
			pt_out^[pos_out] := 109;
			pos_out := pos_out + 1;
			pt_out^[pos_out] := 112;
			pos_out := pos_out + 1;
			pt_out^[pos_out] := 59;
		60: (* < detected *)
			IF pos_out > OSCAT_BASIC.STRING_LENGTH - 4 THEN EXIT; END_IF;
			pt_out^[pos_out] := 38;
			pos_out := pos_out + 1;
			pt_out^[pos_out] := 108;
			pos_out := pos_out + 1;
			pt_out^[pos_out] := 116;
			pos_out := pos_out + 1;
			pt_out^[pos_out] := 59;
		62: (* > detected *)
			IF pos_out > OSCAT_BASIC.STRING_LENGTH - 4 THEN EXIT; END_IF;
			pt_out^[pos_out] := 38;
			pos_out := pos_out + 1;
			pt_out^[pos_out] := 103;
			pos_out := pos_out + 1;
			pt_out^[pos_out] := 116;
			pos_out := pos_out + 1;
			pt_out^[pos_out] := 59;
	ELSE
		IF M AND B > 127 THEN
			tmp := OSCAT_BASIC.CHARNAME(B);
			(* exit if output string has not enough space *)
			IF pos_out + LEN(tmp) + 2 <= 250 THEN
				pt_out^[pos_out] := 38;
				pos_out := pos_out + 1;
				FOR i := 1 TO LEN(tmp) DO
					pt_out^[pos_out] := OSCAT_BASIC.CODE(tmp, i);
					pos_out := pos_out + 1;
				END_FOR;
				pt_out^[pos_out] := 59;
			END_IF;
		ELSE
			pt_out^[pos_out] := B;
		END_IF;
	END_CASE;
	(* increment in by 1 *)
	pos_in := pos_in + 1;
END_FOR;

(* terminate the output string *)
pt_out^[pos_out] := 0;

(* revision history
hm		3. mai. 2008	rev 1.0
	original version

hm		10. mai. 2008	rev 1.1
	stringlength 250
*)
END_FUNCTION

(* ---- HTTP_DEMO.st ---- *)
FUNCTION HTTP_DEMO
VAR
    url_text : STRING := 'http://weather.yahooapis.com/forecastrss?p=94089&u=c';
    URL_DATA : URL;
    IP_C : IP_C;
    S_BUF : NETWORK_BUFFER;
    R_BUF : NETWORK_BUFFER;
    IP_CONTROL_1 : IP_CONTROL;
    DNS_CLIENT : DNS_CLIENT;
    HTTP_GET : HTTP_GET;
    http_release : BOOL;
    enable : BOOL := TRUE;
    http_status : STRING;
    header_start : UINT;
    header_stop : UINT;
    body_start : UINT;
    body_stop : UINT;
    http_get_done : BOOL;
    http_get_error : DWORD;
    COUNT_DR : OSCAT_BASIC.COUNT_DR;
    cycles : DWORD;
    TON_1 : TON;
    F_TRIG : F_TRIG;
END_VAR

END_FUNCTION

(* ---- HYPOT.st ---- *)
FUNCTION HYPOT : REAL
VAR_INPUT
    X : REAL;
    Y : REAL;
END_VAR
HYPOT := SQRT(x*x + y*y);

(* revision history
hm	21. feb 2008	rev 1.0
	original version

*)
END_FUNCTION

(* ---- INC.st ---- *)
FUNCTION INC : INT
VAR_INPUT
    X : INT;
    D : INT;
    M : INT;
END_VAR
INC := (X + D + M + 1) MOD (M + 1);

(* revision history
hm	7. feb 2007		REV 1.0
	original version

hm	15. jan 2008	rev 1.1
	allow for neagtive increment

*)
END_FUNCTION

(* ---- INC1.st ---- *)
FUNCTION INC1 : INT
VAR_INPUT
    X : INT;
    N : INT;
END_VAR
IF X >= N - 1 THEN
	INC1 := 0;
ELSE
	INC1 := X + 1;
END_IF;

(* revision history
hm	13. oct. 2008	rev 1.0
	original version

hm	22. oct. 2008	rev 1.1
	added statement to return value for compatibility reasons

hm	23. feb. 2009	rev 1.2
 	when inc1 is called with X >= N inc will continue with 0
*)
END_FUNCTION

(* ---- INC2.st ---- *)
FUNCTION INC2 : INT
VAR_INPUT
    X : INT;
    D : INT;
    L : INT;
    U : INT;
END_VAR

VAR
    tmp : INT;
END_VAR
tmp := U - L + 1;
INC2 := (X + D - L + tmp) MOD tmp + L;

(* revision history
hm	29. jun. 2008		REV 1.0
	original version

*)
END_FUNCTION

(* ---- INI_PARSER_BUF_DEMO.st ---- *)
FUNCTION INI_PARSER_BUF_DEMO
VAR
    STATION_NAME : STRING;
    STATION_IP : STRING;
    SMTP_SERVER : STRING;
    SMTP_FROM : STRING;
    IPB : INI_PARSER_BUF;
    FS : FILE_SERVER;
    FSD : FILE_SERVER_DATA;
    PT : NETWORK_BUFFER;
    section : INT;
    key : STRING(OSCAT_BASIC.STRING_LENGTH);
    value : STRING(OSCAT_BASIC.STRING_LENGTH);
    str : STRING(OSCAT_BASIC.STRING_LENGTH);
    step : INT;
    result : BYTE;
    offset : UDINT;
    run : BYTE;
    done : BOOL;
END_VAR
(* Demo-Programm: INI-Datei mittels Enumeration auswerten *)

(* ----- den nachfolgenden Textblock als datei "config.ini" auf der sps ablegen ---
# Demo - Initialisierungsdatei

[Station]
NAME=Test_Station_1
IP=192.168.178.1

[SMTP]
SERVER=test.server.de
FROM=test1@gmx.net
---------------------------------------------------------------------------------*)

CASE step OF

00:	IF NOT done THEN
	 	(* File_Daten einrichten  *)
		FSD.FILENAME := 'config.ini'; (* Dateiname *)
		FSD.MODE := 1; (* vorhandene Datei zum lesen öffnen *)
		FSD.OFFSET := 0; (* Start bei Dateianfang *)
		PT.SIZE := 65535; (* maximale länge einlesen *)
		step := 10;
	END_IF;

10:	IF FSD.MODE = 0 THEN (* Datei geöffnet ? *)
		OFFSET := 0; (* Start Offset vorgeben *)
		str := '';
		run := 3; (* key suchen *)
		step := 20;
	END_IF;

20:	IF run = 0 THEN
		(* ---------------------- Debug-Message ----------------------------*)
		(*IF _debug_enable THEN
			LOG_CL.NEW_MSG := 'IPBD: /key >~1< /value >~2< /offset ~3 /Run ~4 /Result ~5';
			LOG_CL.PRINTF[1] := key;
			LOG_CL.PRINTF[2] := value;
			LOG_CL.PRINTF[3] := UDINT_TO_STRING(OFFSET);
			LOG_CL.PRINTF[4] := BYTE_TO_STRING(run);
			LOG_CL.PRINTF[5] := BYTE_TO_STRING(result);
			LOG_MSG();
		END_IF;*)
		(* -----------------------------------------------------------------*)

		run := 3; (* vorbelegung -> naechsten key suchen *)

		IF result = 1 THEN (* neue Sektion gefunden *)
			IF key = 'Station' THEN
				section := 1;
			ELSIF key = 'SMTP' THEN
				section := 2;

			(* hier können weitere Section hinzugefügt werden *)

			ELSE
				section := 0; (* unbekannte sektion gefunden -> ignorieren *)
			END_IF;

		ELSIF result = 2 AND section > 0 THEN (* Key in einer bekannten sektion gefunden *)

			CASE section OF

			1:  (* Section: Station *)
				IF key = 'NAME' THEN
					STATION_NAME := value; (* Name *)
				ELSIF key = 'IP' THEN
					STATION_IP := value; (* IP-Adresse *)
				END_IF;

				(* hier können weitere Schlüsselsauswertungen hinzugefügt werden *)

			2:  (* Section: SMTP *)
				IF key = 'SERVER' THEN
					SMTP_SERVER := value; (* SMTP Server *)
				ELSIF key = 'FROM' THEN
					SMTP_FROM := value; (* SMTP Absender *)
				END_IF;

				(* hier können weitere Schlüsselsauswertungen hinzugefügt werden *)

			END_CASE;

		ELSIF result = 10 THEN (* nichts mehr gefunden *)
			run := 0; (* keine weitere INI Auswertung erwünscht *)
			FSD.MODE := 5; (* Datei schliessen *)
			step := 30;
		END_IF;
	END_IF;

30:	IF FSD.MODE = 0 THEN (* Datei geschlossen ? *)
		step := 0;
		done := TRUE;
	END_IF;

END_CASE;

IPB(STR:=str,RUN:=run,OFFSET:=OFFSET,KEY:=key,VALUE:=value,PT:=PT); (* INI PARAMETER BUF *)
result:=IPB.RESULT;

FS(FSD:=FSD,PT:=PT); (* FILE_SERVER *)
END_FUNCTION

(* ---- INI_PARSER_FILE_DEMO.st ---- *)
FUNCTION INI_PARSER_FILE_DEMO
VAR
    STATION_NAME : STRING;
    STATION_IP : STRING;
    SMTP_SERVER : STRING;
    SMTP_FROM : STRING;
    IPF : INI_PARSER_FILE; // Assuming INI_PARSER_FILE is a previously defined data type
    FS : FILE_SERVER; // Assuming FILE_SERVER is a previously defined data type
    FSD : FILE_SERVER_DATA; // Assuming FILE_SERVER_DATA is a previously defined data type
    PT : NETWORK_BUFFER; // Assuming NETWORK_BUFFER is a previously defined data type
    section : INT;
    filename : STRING;
    key : STRING(OSCAT_BASIC.STRING_LENGTH);
    value : STRING(OSCAT_BASIC.STRING_LENGTH);
    str : STRING(OSCAT_BASIC.STRING_LENGTH);
    step : INT;
    result : BYTE;
    offset : UDINT;
    run : BYTE;
    done : BOOL;
END_VAR
(* Demo-Programm: INI-Datei mittels Enumeration auswerten *)

(* ----- den nachfolgenden Textblock als datei "config.ini" auf der sps ablegen ---
# Demo - Initialisierungsdatei

[Station]
NAME=Test_Station_1
IP=192.168.178.1

[SMTP]
SERVER=test.server.de
FROM=test1@gmx.net
---------------------------------------------------------------------------------*)

CASE step OF

00:	IF NOT done THEN
		filename := 'config.ini'; (* File_Daten einrichten *)
		OFFSET := 0; (* Start Offset vorgeben *)
		str := '';
		run := 3; (* key suchen *)
		step := 20;
	END_IF;

20:	IF run = 0 THEN (* kein Befehl mehr aktiv ? *)
		(* ---------------------- Debug-Message ----------------------------*)
		(*IF _debug_enable THEN
			LOG_CL.NEW_MSG := 'IPFD: /key >~1< /value >~2< /offset ~3 /Run ~4 /Result ~5';
			LOG_CL.PRINTF[1] := key;
			LOG_CL.PRINTF[2] := value;
			LOG_CL.PRINTF[3] := UDINT_TO_STRING(OFFSET);
			LOG_CL.PRINTF[4] := BYTE_TO_STRING(run);
			LOG_CL.PRINTF[5] := BYTE_TO_STRING(result);
			LOG_MSG();
		END_IF;*)
		(* -----------------------------------------------------------------*)

		run := 3; (* vorbelegung -> naechsten key suchen *)

		IF result = 1 THEN (* neue Sektion gefunden *)
			IF key = 'Station' THEN
				section := 1;
			ELSIF key = 'SMTP' THEN
				section := 2;

			(* hier können weitere Section hinzugefügt werden *)

			ELSE
				section := 0; (* unbekannte sektion gefunden -> ignorieren *)
			END_IF;

		ELSIF result = 2 AND section > 0 THEN (* Key in einer bekannten sektion gefunden *)

			CASE section OF

			1:  (* Section: Station *)
				IF key = 'NAME' THEN
					STATION_NAME := value; (* Name *)
				ELSIF key = 'IP' THEN
					STATION_IP := value; (* IP-Adresse *)
				END_IF;

				(* hier können weitere Schlüsselsauswertungen hinzugefügt werden *)

			2:  (* Section: SMTP *)
				IF key = 'SERVER' THEN
					SMTP_SERVER := value; (* SMTP Server *)
				ELSIF key = 'FROM' THEN
					SMTP_FROM := value; (* SMTP Absender *)
				END_IF;

				(* hier können weitere Schlüsselsauswertungen hinzugefügt werden *)

			END_CASE;

		ELSIF result = 10 THEN (* nichts mehr gefunden *)
			run := 0; (* keine weitere INI Auswertung erwünscht *)
			FSD.MODE := 5; (* Datei schliessen *)
			step := 30;
		END_IF;
	END_IF;

30:	IF FSD.MODE = 0 THEN (* Befehl Datei schliessen beendet *)
		step := 0;
		done := TRUE;
	END_IF;

END_CASE;

IPF(FILENAME:=FILENAME,FSD:=FSD,STR:=str,RUN:=run,OFFSET:=OFFSET,KEY:=key,VALUE:=value,PT:=PT); (* INI PARAMETER FILE *)
result:=IPF.RESULT;

FS(FSD:=FSD,PT:=PT); (* FILE_SERVER *)
END_FUNCTION

(* ---- INT_TO_BCDC.st ---- *)
FUNCTION INT_TO_BCDC : BYTE
VAR_INPUT
    IN : INT;
END_VAR
INT_TO_BCDC := SHL(INT_TO_BYTE(IN / INT#10),4) OR INT_TO_BYTE(in MOD INT#10);

(* revision history
hm	13.12.2007
	original version

hm	30.6.2008	rev 1.1
	changed name INT_TO_BCD to INT_TO_BCDC to avoid collision with util.lib
	corrected error in code

*)
END_FUNCTION

(* ---- INV.st ---- *)
FUNCTION INV : REAL
VAR_INPUT
    X : REAL;
END_VAR
IF X <> 0.0 THEN INV := 1.0 / X; END_IF;

(* revision history
hm	26. oct. 2008	rev 1.0
	original version

hm	10. mar. 2009	rev 1.1
	real constants updated to new systax using dot

*)
END_FUNCTION

(* ---- IP2GEO_DEMO.st ---- *)
FUNCTION IP2GEO_DEMO
VAR
    IP_C : IP_C;
    S_BUF : NETWORK_BUFFER;
    R_BUF : NETWORK_BUFFER;
    IP_CONTROL_1 : IP_CONTROL;
    CLK_PRG : oscat_basic.CLK_PRG;
    IP2GEO_1 : IP2GEO;
    GEO : IP2GEO_DATA;
    activate : BOOL := TRUE;
    done : BOOL;
    busy : BOOL;
    error_c : DWORD;
    error_t : BYTE;
END_VAR

END_FUNCTION

(* ---- IP4_CHECK.st ---- *)
FUNCTION IP4_CHECK : BOOL
VAR_INPUT
    NIP : DWORD;
    LIP : DWORD;
    SM  : DWORD;
END_VAR
IP4_CHECK := (NIP AND sm) = (LIP AND SM);

(* revision history
hm		4. mar 2008	rev 1.0
	original version

*)
END_FUNCTION

(* ---- IP4_DECODE.st ---- *)
FUNCTION IP4_DECODE : DWORD
VAR_INPUT
    str : STRING(15);
END_VAR

VAR
    pos : INT;
END_VAR
pos := FIND(str, '.');
WHILE pos > 0 DO
	IP4_DECODE := SHL(IP4_DECODE,8) OR STRING_TO_DWORD(LEFT(str,pos - 1));
	str := DELETE(str, pos, 1);
	pos := FIND(str, '.');
END_WHILE;
IP4_DECODE := SHL(IP4_DECODE,8) OR STRING_TO_DWORD(str);

(* revision history
hm		29. feb 2008	rev 1.0
	original version

hm	10. mar. 2009	rev 1.1
	new algorythm
*)
END_FUNCTION

(* ---- IP4_TO_STRING.st ---- *)
FUNCTION IP4_TO_STRING : string
VAR_INPUT
    IP4 : DWORD;
END_VAR

VAR
    tmp : STRING[3];
END_VAR
(* mask bits AND INSERT AT given position *)
tmp := BYTE_TO_STRING(DWORD_TO_BYTE(IP4));
IP4_TO_STRING := CONCAT('...', tmp);
tmp := BYTE_TO_STRING(DWORD_TO_BYTE(SHR(IP4,8)));
IP4_TO_STRING := INSERT(IP4_TO_STRING, tmp, 2);
tmp := BYTE_TO_STRING(DWORD_TO_BYTE(SHR(IP4,16)));
IP4_TO_STRING := INSERT(IP4_TO_STRING, tmp, 1);
tmp := BYTE_TO_STRING(DWORD_TO_BYTE(SHR(IP4,24)));
IP4_TO_STRING := CONCAT(tmp, IP4_TO_STRING);

(* revision history
hm	22. apr 2008	rev 1.0
	original version

hm	10. mar. 2009	rev 1.1
	improved code
*)
END_FUNCTION

(* ---- IRTRANS_DEMO.st ---- *)
FUNCTION IRTRANS_DEMO
VAR
    IP_C : IP_C;
    S_BUF : NETWORK_BUFFER_SHORT;
    R_BUF : NETWORK_BUFFER_SHORT;
    IP_CONTROL2 : IP_CONTROL2;
    IRTRANS_DECODE : IRTRANS_DECODE;
    IRTRANS_RCV_4 : IRTRANS_RCV_4;
    DRIVER_4 : oscat_basic.DRIVER_4;
    IRTRANS_SERVER : IRTRANS_SERVER;
    IRTRANS_SND_8_1 : IRTRANS_SND_8;
    IRTRANS_SND_8_2 : IRTRANS_SND_8;
    Q0 : BOOL;
    Q1 : BOOL;
    Q2 : BOOL;
    Q3 : BOOL;
    error : BOOL;
    error_server : DWORD;
    Send_1_0 : BOOL := TRUE;
    Send_1_1 : BOOL;
    Send_1_2 : BOOL;
    Send_1_3 : BOOL;
    Send_1_4 : BOOL;
    Send_1_5 : BOOL;
    Send_1_6 : BOOL;
    Send_1_7 : BOOL;
    Send_2_0 : BOOL := TRUE;
    Send_2_1 : BOOL;
    Send_2_2 : BOOL;
    Send_2_3 : BOOL;
    Send_2_4 : BOOL;
    Send_2_5 : BOOL;
    Send_2_6 : BOOL;
    Send_2_7 : BOOL;
    R_ENABLE : BOOL;
    S_ENABLE : BOOL;
    MODE : BOOL := FALSE;
    KEY_1 : BYTE;
    KEY_2 : BYTE;
END_VAR

END_FUNCTION

(* ---- IS_ALNUM.st ---- *)
FUNCTION IS_ALNUM : BOOL
VAR_INPUT
    str : STRING(STRING_LENGTH);
END_VAR_INPUT

VAR
    L : INT;
    pt : POINTER TO BYTE;
    pos : INT;
END_VAR
PT := ADR(str);
L := LEN(str);
FOR pos := 1 TO L DO
	IF NOT (ISC_ALPHA(pt^) OR ISC_NUM(pt^)) THEN
		IS_ALNUM := FALSE;
		RETURN;
	END_IF;
    	PT := PT + 1;
END_FOR;
IS_ALNUM := L > 0;

(* revision history
hm	29. feb 2008	rev 1.0
	original version

hm	29. mar. 2008	rev 1.1
	changed STRING to STRING(STRING_LENGTH)
*)
END_FUNCTION

(* ---- IS_ALPHA.st ---- *)
FUNCTION IS_ALPHA : BOOL
VAR_INPUT
    str: STRING(STRING_LENGTH);
END_VAR

VAR
    L: INT;
    pt: POINTER TO BYTE;
    pos: INT;
END_VAR
PT := ADR(str);
L := LEN(str);
FOR pos := 1 TO L DO
	IF NOT ISC_ALPHA(pt^) THEN
		IS_ALPHA := FALSE;
		RETURN;
	END_IF;
    	PT := PT + 1;
END_FOR;
IS_ALPHA := L > 0;

(* revision history
hm	29. feb 2008	rev 1.0
	original version

hm	29. mar. 2008	rev 1.1
	changed STRING to STRING(STRING_LENGTH)
*)
END_FUNCTION

(* ---- IS_CC.st ---- *)
FUNCTION IS_CC : BOOL
VAR_INPUT
    str : STRING(STRING_LENGTH);
    cmp : STRING(STRING_LENGTH);
END_VAR

VAR
    L : INT;
    pos : INT;
END_VAR
L := LEN(str);
FOR pos := 1 TO L DO
	IF FIND(CMP,MID(str,1,pos)) = 0 THEN RETURN; END_IF;
END_FOR;
IS_CC := L > 0;

(* revision history
hm	19. mar 2008	rev 1.0
	original version

hm	29. mar. 2008	rev 1.1
	changed STRING to STRING(STRING_LENGTH)
*)
END_FUNCTION

(* ---- IS_CTRL.st ---- *)
FUNCTION IS_CTRL : BOOL
VAR_INPUT
    STR : STRING(STRING_LENGTH);
END_VAR

VAR
    L : INT;
    pt : POINTER TO BYTE;
    pos : INT;
END_VAR
PT := ADR(str);
L := LEN(str);
FOR pos := 1 TO L DO
	IF NOT (ISC_CTRL(pt^)) THEN
		IS_CTRL := FALSE;
		RETURN;
	END_IF;
    	PT := PT + 1;
END_FOR;
IS_CTRL := L > 0;

(* revision history
hm	29. feb. 2008	rev 1.0
	original version

hm	29. mar. 2008	rev 1.1
	changed STRING to STRING(STRING_LENGTH)
*)
END_FUNCTION

(* ---- IS_HEX.st ---- *)
FUNCTION IS_HEX : BOOL
VAR_INPUT
    str : STRING[STRING_LENGTH];
END_VAR

VAR
    L : INT;
    pt : POINTER TO BYTE;
    pos : INT;
END_VAR
PT := ADR(str);
L := LEN(str);
FOR pos := 1 TO L DO
	IF NOT (ISC_HEX(pt^)) THEN
		IS_HEX := FALSE;
		RETURN;
	END_IF;
    	PT := PT + 1;
END_FOR;
IS_HEX := L > 0;

(* revision history
hm	29. feb 2008	rev 1.0
	original version

hm	29. mar. 2008	rev 1.1
	changed STRING to STRING(STRING_LENGTH)
*)
END_FUNCTION

(* ---- IS_IP4.st ---- *)
FUNCTION IS_IP4 : BOOL
VAR_INPUT
    str : STRING;
END_VAR
IS_IP4 := OSCAT_BASIC.COUNT_CHAR(str, 46) = 3;

(* revision history
hm	1. mar. 2008	rev 1.0
	original version

hm	10. mar. 2009	rev 1.1
	new code

*)
END_FUNCTION

(* ---- IS_LOWER.st ---- *)
FUNCTION IS_LOWER : BOOL
VAR_INPUT
    str : STRING[STRING_LENGTH]; // Input variable declaration
END_VAR

VAR
    l : INT; // Local variable declaration
    pt : POINTER TO BYTE; // Pointer variable declaration
    pos : INT; // Position variable declaration
END_VAR
PT := ADR(str);
L := LEN(str);
FOR pos := 1 TO L DO
	IF NOT (ISC_LOWER(pt^)) THEN
		IS_LOWER := FALSE;
		RETURN;
	END_IF;
    	PT := PT + 1;
END_FOR;
IS_LOWER := L > 0;

(* revision history
hm	29. feb 2008	rev 1.0
	original version

hm	29. mar. 2008	rev 1.1
	changed STRING to STRING(STRING_LENGTH)
*)
END_FUNCTION

(* ---- IS_NCC.st ---- *)
FUNCTION IS_NCC : BOOL
VAR_INPUT
    str : STRING[STRING_LENGTH];
    cmp : STRING[STRING_LENGTH];
END_VAR

VAR
    L : INT;
    pos : INT;
END_VAR
L := LEN(str);
FOR pos := 1 TO L DO
	IF FIND(CMP,MID(str,1,pos)) > 0 THEN RETURN; END_IF;
END_FOR;
IS_NCC := TRUE;

(* revision history
hm	19. mar 2008	rev 1.0
	original version

hm	29. mar. 2008	rev 1.1
	changed STRING to STRING(STRING_LENGTH)
*)
END_FUNCTION

(* ---- IS_NUM.st ---- *)
FUNCTION IS_NUM : BOOL
VAR_INPUT
    str : STRING[STRING_LENGTH];  // Input variable of type STRING with specified length
END_VAR

VAR
    L : INT;                       // Local variable of type INT
    pt : POINTER TO BYTE;         // Local variable, pointer to BYTE
    pos : INT;                    // Local variable of type INT
END_VAR
PT := ADR(str);
L := LEN(str);
FOR pos := 1 TO L DO
	IF NOT (ISC_NUM(pt^)) THEN
		IS_NUM := FALSE;
		RETURN;
	END_IF;
    	PT := PT + 1;
END_FOR;
IS_NUM := L > 0;

(* revision history
hm	29. feb 2008	rev 1.0
	original version

hm	29. mar. 2008	rev 1.1
	changed STRING to STRING(STRING_LENGTH)
*)
END_FUNCTION

(* ---- IS_SORTED.st ---- *)
FUNCTION IS_SORTED : BOOL
VAR_INPUT
    pt : ^ ARRAY [0..32000] OF REAL; // Pointer to an array of REAL
    size : UINT; // Size variable of type UINT
END_VAR

VAR
    stop : INT; // Local variable of type INT
    i : INT; // Local variable of type INT
END_VAR
stop := UINT_TO_INT(SHR(size,2)-2);
FOR i := 0 TO stop DO
	IF pt^[i] > pt^[i+1] THEN
		IS_SORTED := FALSE;
		RETURN;
	END_IF;
END_FOR;

IS_SORTED := TRUE;

(* revision history

hm 	29. mar. 2008 	rev 1.0
	original version

hm	4. apr. 2008	rev 1.1
	added type conversion to avoid warnings under codesys 3.0
*)
END_FUNCTION

(* ---- IS_UPPER.st ---- *)
FUNCTION IS_UPPER : BOOL
VAR_INPUT
    str : STRING; // Length to be defined as per application requirements
END_VAR

VAR
    L : INT;
    pt : POINTER TO BYTE;
    pos : INT;
END_VAR
PT := ADR(str);
L := LEN(str);
FOR pos := 1 TO L DO
	IF NOT (ISC_UPPER(pt^)) THEN
		IS_UPPER := FALSE;
		RETURN;
	END_IF;
    	PT := PT + 1;
END_FOR;
IS_UPPER := L > 0;

(* revision history
hm	29. feb 2008	rev 1.0
	original version

hm	29. mar. 2008	rev 1.1
	changed STRING to STRING(STRING_LENGTH)
*)
END_FUNCTION

(* ---- IS_URLCHR.st ---- *)
FUNCTION IS_URLCHR : BOOL
VAR_INPUT
    IN : BYTE;
END_VAR
IS_URLCHR := ((IN > 47) AND (IN < 58)) OR ((IN > 64) AND (IN < 91)) OR ((IN > 96) AND (IN < 123)) OR (in = 126) OR (in = 95) OR (in =45) OR (in =46);

(* revision history
hm		27. apr. 2008	rev 1.0
	original version

*)
END_FUNCTION

(* ---- ISC_ALPHA.st ---- *)
FUNCTION ISC_ALPHA : BOOL
#VAR_INPUT
    IN : BYTE;
END_VAR
IF setup.EXTENDED_ASCII THEN
	ISC_ALPHA := (in > 64 AND in < 91) OR (in > 191  AND in <> 215 AND in <> 247) OR (in > 96 AND in < 123);
ELSE
	ISC_ALPHA := (IN > 64 AND IN < 91) OR (in > 96 AND in < 123);
END_IF;

(* revision history
hm	6. mar. 2008	rev 1.0
	original version

hm	19. oct. 2008	rev 1.1
	changes setup constants
*)
END_FUNCTION

(* ---- ISC_CTRL.st ---- *)
FUNCTION ISC_CTRL : BOOL
VAR_INPUT
    IN : BYTE;
END_VAR
ISC_CTRL := IN < 32 OR IN = 127;

(* revision history
hm		6. mar. 2008	rev 1.0
	original version

*)
END_FUNCTION

(* ---- ISC_HEX.st ---- *)
FUNCTION ISC_HEX : BOOL
VAR_INPUT
    IN : BYTE;
END_VAR
ISC_HEX := (IN > 47 AND IN < 58) OR (IN > 64 AND IN < 71) OR (IN > 96 AND IN < 103);

(* revision history
hm		6. mar. 2008	rev 1.0
	original version

*)
END_FUNCTION

(* ---- ISC_LOWER.st ---- *)
FUNCTION ISC_LOWER : BOOL
VAR_INPUT
    IN : BYTE; // Input variable
END_VAR
IF setup.EXTENDED_ASCII THEN
	ISC_LOWER := ((in > 96) AND (in < 123)) OR ((in > 222) AND (in <> 247));
ELSE
	ISC_LOWER := ((in > 96) AND (in < 123));
END_IF;

(* revision history
hm	6. mar. 2008	rev 1.0
	original version

hm	19. oct. 2008	rev 1.1
	changes setup constants
*)
END_FUNCTION

(* ---- ISC_NUM.st ---- *)
FUNCTION ISC_NUM : BOOL
VAR_INPUT
    IN : BYTE;
END_VAR
ISC_NUM := IN > 47 AND IN < 58;

(* revision history
hm		6. mar. 2008	rev 1.0
	original version

*)
END_FUNCTION

(* ---- ISC_UPPER.st ---- *)
FUNCTION ISC_UPPER : BOOL
VAR_INPUT
    IN : BYTE;
END_VAR
IF setup.EXTENDED_ASCII THEN
	ISC_UPPER :=  ((in > 64) AND (in < 91)) OR (((in > 191) AND (in < 223)) AND (in <> 215));
ELSE
	ISC_UPPER := ((in > 64) AND (in < 91));
END_IF;

(* revision history
hm	6. mar. 2008	rev 1.0
	original version

hm	19. oct. 2008	rev 1.1
	changes setup constants

*)
END_FUNCTION

(* ---- JD2000.st ---- *)
FUNCTION JD2000 : REAL
VAR_INPUT
    DTI : TIME;
END_VAR
JD2000 := DWORD_TO_REAL(DT_TO_DWORD(DTI) - 946728000) / 86400.0;

(* revision histroy
hm	15. jul. 2008	rev 1.0
	original release

*)
END_FUNCTION

(* ---- K_TO_C.st ---- *)
FUNCTION K_TO_C : REAL
VAR_INPUT
    Kelvin : REAL;
END_VAR
K_TO_C := Kelvin + phys.T0;

(* revision history

hm	4. aug 2006	rev 1.0
	original version

hm	19. aug 2009	rev 1.1
	fixed calculation error

*)
END_FUNCTION

(* ---- KMH_TO_MS.st ---- *)
FUNCTION KMH_TO_MS : REAL
VAR_INPUT
    kmh : REAL;
END_VAR
KMH_TO_MS := kmh * 0.2777777777777;

(* revision history
hm	4. feb 2007		rev 1.0
	original version

hm	6. jan 2008		rev 1.1
	improved performance

*)
END_FUNCTION

(* ---- LAMBERT_W.st ---- *)
FUNCTION LAMBERT_W : REAL
VAR_INPUT
    X : REAL;
END_VAR

VAR
    w : REAL;
    i : INT;
    we : REAL;
    w1e : REAL;
    last : DWORD;
    ewx : REAL;
END_VAR
(* check for valid input and return -1000 if too low *)
IF x < -0.367879441171442 THEN
	LAMBERT_W := -1000.0;
	RETURN;
(* return 0 if x = 0 *)
ELSIF x = 0.0 THEN
	RETURN;
(* first an estimate is calculated *)
ELSIF x <= 500.0 THEN
	w := LN(x + 1.0);
	w := 0.665 * (1.0 + 0.0195 * w) * w + 0.04;
ELSE
	w := LN(x - 4.0) - (1.0 - 1.0/LN(x)) * LN(LN(x));
END_IF;
(* use estimate to calculate exact result *)
FOR i := 0 TO 5 DO
	ewx := EXP(w);
	we := w * ewx - x;
	w1e := (w+1.0) * ewx;
	last := REAL_TO_DW(w) AND 16#FFFF_FFFC;
	w := w - (we / (w1e - (w+2.0) * we / (2.0 * w + 2.0)));
	IF (REAL_TO_DW(w) AND 16#FFFF_FFFC) = last THEN EXIT; END_IF;
END_FOR;
LAMBERT_W := w;

(* revision hisdtory
hm	26. oct. 2008	rev 1.0
	original version

hm	10. mar. 2009	rev 1.1
	real constants updated to new systax using dot

*)
END_FUNCTION

(* ---- LANGEVIN.st ---- *)
FUNCTION LANGEVIN : REAL
VAR_INPUT
    X : REAL;
END_VAR
IF X = 0.0 THEN
	LANGEVIN := 0.0;
ELSE
	LANGEVIN := COTH(X) - 1.0 / X;
END_IF;

(* revision history
hm	10.12.2007	rev 1.0
	original version

hm	11. mar 2008	rev 1.1
	changed formula to avoid problems when x = 0

hm	10. mar. 2009	rev 1.2
	real constants updated to new systax using dot

*)
END_FUNCTION

(* ---- LEAP_DAY.st ---- *)
FUNCTION LEAP_DAY : BOOL
VAR_INPUT
    IDATE : DATE;
END_VAR
LEAP_DAY := DATE_TO_UDINT(IDATE) MOD 126230400 = 68169600;

(* change history

hm 	15. jun. 2008	rev 1.0
	original version

hm	7. oct. 2008	rev 1.1
	changed function month to month_of_date

hm	24. jan. 2011	rev 1.2
	improved performance
*)
END_FUNCTION

(* ---- LEAP_OF_DATE.st ---- *)
FUNCTION LEAP_OF_DATE : BOOL
VAR_INPUT
    idate: DATE;
END_VAR
LEAP_OF_DATE := SHL(((DATE_TO_DWORD(idate) + 43200) / 31557600), 30) = 16#80000000;

(* change history

2.10.2006		rev 1.1
the function now calls leap_year to accomodate further accuracy.
the function now works for any year from 1970 to 2100

8. jan 2008		rev 1.2
	improved code for better performance

28. jan. 2011	rev 1.3
	improved performance
*)
END_FUNCTION

(* ---- LEAP_YEAR.st ---- *)
FUNCTION LEAP_YEAR : BOOL
VAR_INPUT
    yr : INT;  // Variable for year
END_VAR
LEAP_YEAR := SHL(yr,14) = 0;

(* this code was used prior to rev 1.1

IF yr MOD 400 = 0 THEN leap_year := TRUE;
ELSIF yr MOD 100 = 0 THEN leap_year := FALSE;
ELSIF yr MOD 4 =0 THEN leap_year := TRUE;
ELSE leap_year := FALSE;
END_IF;

*)

(* change history

hm 	2.10.2006		rev 1.1
	the function now works for any year from 1970 up to 2100

hm	1. oct 2007		rev 1.2
	chaged code for higher performance
*)
END_FUNCTION

(* ---- LINEAR_INT.st ---- *)
FUNCTION LINEAR_INT : REAL
VAR_INPUT
    X : REAL;
    XY : ARRAY[1..20, 0..1] OF REAL;
    Pts : INT;
END_VAR

VAR
    i : INT;
END_VAR
(*make sure n is bound within the array size *)
pts := MIN(pts,20);

(* calculate the linear segement interpolation *)
i := 2;
(* search for segment and calculate output
	below and above the defined segments we interpolate the last segment *)
WHILE (i < pts) AND (XY[i,0] < X) DO
	i := i + 1;
END_WHILE;

(* calculate the output value on the corresponding segment coordinates *)
LINEAR_INT := ((XY[i,1] - XY[i-1,1]) * X - XY[i,1] * XY[i-1,0] + XY[i-1,1] * XY[i,0]) / (XY[i,0] - XY[i-1,0]);

(* revision history
hm	7. oct 2007		rev 1.0
	original version

hm	27 dec 2007		rev 1.1
	changed code for better performance
*)
END_FUNCTION

(* ---- LIST_ADD.st ---- *)
FUNCTION LIST_ADD : BOOL
VAR_INPUT
    SEP : BYTE;
    INS : STRING(LIST_LENGTH);
END_VAR

VAR_IN_OUT
    LIST : STRING(LIST_LENGTH);
END_VAR

VAR
    sx : STRING(1);
END_VAR
sx := CHR_TO_STRING(SEP);			(* convert separation character to string *)
INS := CONCAT(sx, INS);					(* start element with separation character *)

IF LEN(LIST) + LEN(INS) > LIST_LENGTH THEN
	LIST_ADD := FALSE;					(* return false if element does not fit *)
ELSE
	LIST := CONCAT(LIST, INS);
	LIST_ADD := TRUE;
END_IF;

(* revision histroy

hm	21. mar. 2011	rev 2.0
	original release
*)
END_FUNCTION

(* ---- LIST_CLEAN.st ---- *)
FUNCTION LIST_CLEAN : BOOL
VAR_INPUT
    SEP : BYTE;
END_VAR

VAR_IN_OUT
    LIST : STRING[LIST_LENGTH];
END_VAR

VAR
    pt : POINTER TO ARRAY[1..LIST_LENGTH] OF BYTE;
    read : INT := 1;
    write : INT := 1;
    last : BYTE;
    c : BYTE;
END_VAR
pt := ADR(LIST);

FOR read := 1 TO LIST_LENGTH DO
	c := pt^[read];								(* read character from list *)
	IF c = 0 THEN EXIT;						(* exit the loop if character definbes end of string *)
	ELSIF c <> SEP OR sep <> last THEN	(* copy element from read to write position unless a double sep character is present *)
		pt^[write] := c;
		write := write + 1;
	END_IF;
	last := c;									(* remember last character *)
END_FOR;

IF last = SEP THEN write := write - 1; END_IF;		(* if last character is sep then delete empty element at end *)
IF write <= STRING_LENGTH THEN pt^[write] := 0;	 END_IF;		(* terminate string with 0 *)

LIST_CLEAN := TRUE;						(* retrun TRUE *)

(* revision histroy
hm	28. jun. 2008	rev 1.0
	original release

hm	19. jan. 2011	rev 1.1
	changed string(255) to string(LIST_LENGTH)

hm	21. mar. 2011	rev 2.0
	all elements start with SEP

*)
END_FUNCTION

(* ---- LIST_GET.st ---- *)
FUNCTION LIST_GET : string
VAR_INPUT
    SEP : BYTE;       // Input variable
    POS : INT;        // Input variable
END_VAR

VAR_IN_OUT
    LIST : STRING(LIST_LENGTH);  // InOut variable
END_VAR

VAR
    i : INT := 1;      // Local variable with initial value
    o : INT := 1;      // Local variable with initial value
    pt : POINTER TO ARRAY[1..LIST_LENGTH] OF BYTE; // Pointer to array of BYTE
    po : POINTER TO ARRAY[1..LIST_LENGTH] OF BYTE; // Pointer to array of BYTE
    cnt : INT := 0;    // Local variable with initial value
    c : BYTE;          // Local variable
END_VAR
pt := ADR(LIST);							(* load pointers *)
po := ADR(LIST_GET);

REPEAT
	c := pt^[i];
	IF cnt = pos THEN						(* copy element to output string *)
		IF c = SEP  THEN EXIT; END_IF;		(* next element stop copy and finish *)
		po^[o] := c;
		o := o + 1;
	ELSIF c = SEP THEN
		cnt := cnt + 1;
	END_IF;
	i := i + 1;
UNTIL
	(i = LIST_LENGTH) OR (c = 0)
END_REPEAT;
po^[o] := 0;						(* close the output string *)

(* revision histroy
hm	20. jun. 2008	rev 1.0
	original release

hm	19. jan. 2011	rev 1.1
	changed string(255) to strring(LIST_LENGTH)

hm	21. mar. 2011	rev 2.0
	all list elements start with SEP
*)
END_FUNCTION

(* ---- LIST_INSERT.st ---- *)
FUNCTION LIST_INSERT : BOOL
VAR_INPUT
    SEP : BYTE;
    POS : INT;
    INS : STRING(LIST_LENGTH);
END_VAR

VAR_IN_OUT
    LIST : STRING(LIST_LENGTH);
END_VAR

VAR
    pt : POINTER TO ARRAY[1..LIST_LENGTH] OF BYTE;
    read : INT := 1;
    cnt : INT := 1;
    sx : STRING(1);
END_VAR
(* load pointers *)
pt := ADR(LIST);

IF LEN(ins) + 1 + LEN(LIST) > LIST_LENGTH THEN
	LIST_INSERT := FALSE;
ELSE
	LIST_INSERT := TRUE;
	(* search for position *)
	WHILE read < LIST_LENGTH DO
		IF cnt >= POS THEN
			sx := CHR_TO_STRING(SEP);
			INS := CONCAT(sx, INS);
			LIST := INSERT(LIST, INS, read - 1);
			LIST_INSERT := TRUE;
			RETURN;
		END_IF;
		IF pt^[read]  = 0 THEN				(* list is too short add empty element *)
			pt^[read] := SEP;
			pt^[read + 1] := 0;
		END_IF;
		read := read + 1;
		IF pt^[read] = SEP OR pt^[read] = 0 THEN cnt := cnt + 1; END_IF;
	END_WHILE;
END_IF;

(* revision histroy
hm	28. jun. 2008	rev 1.0
	original release

hm	17. dec. 2008	rev 1.1
	changes name of function chr to chr_to_string

hm	19. jan. 2011	rev 1.2
	changed string(255) to string(LIST_LENGTH)

hm	21. mar. 2011	rev 2.0
	all list elements start with SEP

*)
END_FUNCTION

(* ---- LIST_LEN.st ---- *)
FUNCTION LIST_LEN : INT
VAR_INPUT
    SEP : BYTE;
END_VAR

VAR_IN_OUT
    LIST : STRING(LIST_LENGTH);
END_VAR

VAR
    pt : ^ARRAY[1..LIST_LENGTH] OF BYTE;
    pos : INT := 1;
    c : BYTE;
END_VAR
pt := ADR(LIST);
LIST_LEN := 0;
REPEAT
	c := pt^[pos];
	IF c = SEP THEN LIST_LEN := LIST_LEN + 1; END_IF;
	pos := pos + 1;
UNTIL
	c = 0 OR pos > LIST_LENGTH
END_REPEAT;

(* revision histroy
hm	25. jun. 2008	rev 1.0
	original release

hm	16. oct. 2008	rev 1.1
	fixed a problem where list_len would only work up to LIST_LENGTH

hm	19. jan. 2001	rev 1.2
	changed string(255) to string(LIST_LENGTH)

hm	21. mar. 2011	rev 2.0
	all list elements start with SEP

*)
END_FUNCTION

(* ---- LIST_RETRIEVE.st ---- *)
FUNCTION LIST_RETRIEVE : string
VAR_INPUT
    SEP : BYTE;
    POS : INT;
END_VAR

VAR_IN_OUT
    LIST : STRING(LIST_LENGTH);
END_VAR

VAR
    i : INT;
    o : INT := 1;
    w : INT := 1;
    pt : POINTER TO ARRAY[1..LIST_LENGTH] OF BYTE;
    po : POINTER TO ARRAY[1..LIST_LENGTH] OF BYTE;
    cnt : INT := 0;
    c : BYTE;
END_VAR
(* load pointers *)
pt := ADR(LIST);
po := ADR(LIST_RETRIEVE);

IF pos > 0 THEN
	FOR i := 1 TO LIST_LENGTH DO
		c := pt^[i];
		IF c = 0 THEN
			po^[o] := 0;
			IF cnt < pos THEN pt^[w + 1] := 0; ELSE pt^[w] := 0; END_IF;
			RETURN;
		ELSIF cnt = pos AND c <> SEP THEN				(* we have found the element *)
			po^[o] := pt^[i];
			o := o + 1;
		ELSIF cnt >= pos THEN
			pt^[w] := c;
			w := w + 1;
		ELSE
			w := i;
		END_IF;
		IF c = sep THEN cnt := cnt + 1; END_IF;
	END_FOR;
ELSE
	LIST_RETRIEVE := '';
END_IF;

(* revision histroy
hm	28. jun. 2008	rev 1.0
	original release

hm	19. jan. 2011	rev 1.1
	changed string(255) to string(LIST_LENGTH)

hm	21. mar. 2011	rev 2.0
	all elements start with SEP
*)
END_FUNCTION

(* ---- LIST_RETRIEVE_LAST.st ---- *)
FUNCTION LIST_RETRIEVE_LAST : string
VAR_INPUT
    SEP : BYTE;
END_VAR

VAR_IN_OUT
    LIST : STRING[LENGTH := LIST_LENGTH];
END_VAR

VAR
    i : INT;
    last : INT := 1;
    pt : POINTER TO ARRAY[1..LIST_LENGTH] OF BYTE;
    c : BYTE;
END_VAR
(* load pointers *)
pt := ADR(LIST);

(* search position of last element *)
FOR i := 1 TO LIST_LENGTH DO
	c := pt^[i];
	IF c = 0 THEN
		EXIT;
	ELSIF C = SEP THEN
		last := i;
	END_IF;
END_FOR;
(* return last element of list *)
LIST_RETRIEVE_LAST := MID(LIST, LIST_LENGTH, last + 1);
(* terminate list at i *)
pt^[last] := 0;

(* revision histroy
hm	21. mar. 2011	rev 2.0
	new module
*)
END_FUNCTION

(* ---- LOWERCASE.st ---- *)
FUNCTION LOWERCASE : string
VAR_INPUT
    str: STRING[STRING_LENGTH];
END_VAR

VAR
    PT: POINTER TO BYTE;
    pos: INT;
    l: INT;
END_VAR
PT := ADR(LOWERCASE);
lowercase := str;
l := LEN(str);
FOR pos := 1 TO l DO
	pt^ := TO_LOWER(pt^);
	PT := PT + 1;
END_FOR;

(* revision histroy
hm	6. oct. 2006	rev 1.0
	original release

hm	4. feb. 2008	rev 1.1
	improved performance
	added Ä.Ö,Ü

hm	6. mar. 2008	rev 1.2
	added support for exteded Ascii

hm	29. mar. 2008	rev 1.3
	changed STRING to STRING(STRING_LENGTH)
*)
END_FUNCTION

(* ---- LTIME_TO_UTC.st ---- *)
FUNCTION LTIME_TO_UTC : DT
VAR_INPUT
    LOCAL_TIME : DT;
    DST : BOOL;
    TIME_ZONE_OFFSET : INT;
END_VAR
LTIME_TO_UTC := UDINT_TO_DT(DT_TO_UDINT(LOCAL_TIME) - INT_TO_UDINT(TIME_ZONE_OFFSET) * 60);
IF DST THEN LTIME_TO_UTC := LTIME_TO_UTC - T#1h; END_IF;

(* revision history
hm 5.7.2007		rev 1.0
	original version

hm 5.11.2007		rev 1.1
	replaced literal constant with variable because of error in möller ecp4 compiler

hm	12.nov 2007	rev 1.2
	changed Type of time_zone_offset from time to int to allow for time zones with negative offset

hm	8. dec 2007	rev 1.3
	corrected a problem with time_zone_offset

hm	14. oct. 2008	rev 1.4
	changed time_zone_offset from int to real to allow for half hour offset

hm	20. oct. 2006	rev 1.5
	changed time_zone_offset from Real to INT, now in Minutes

hm	27. feb. 2009	rev 1.6
	added type conversions to avoid warnings under codesys 3.0

ks	13. nov. 2009	rev 1.7
	corrected error in formula

*)
END_FUNCTION

(* ---- MANUAL.st ---- *)
FUNCTION MANUAL : BOOL
VAR_INPUT
    IN : BOOL;
    ON : BOOL;
    OFF : BOOL;
END_VAR
MANUAL := NOT OFF AND (IN OR ON);

(* revision history
hm	21. nov 2008	rev 1.0
	original version

*)
END_FUNCTION

(* ---- MAX3.st ---- *)
FUNCTION MAX3 : REAL
VAR_INPUT
    in1 : REAL;
    in2 : REAL;
    in3 : REAL;
END_VAR
MAX3 := MAX(MAX(IN1,IN2),IN3);

(* revision history
hm	1.1.2007	rev 1.0
	original release

hm	18. mar. 2011	rev 1.1
	improve performance

*)
END_FUNCTION

(* ---- MB_CLIENT_DEMO.st ---- *)
FUNCTION MB_CLIENT_DEMO
VAR
    IP_CONTROL2_1 : IP_CONTROL2;
    MB_CLIENT_1 : MB_CLIENT;
    IP_C : IP_C;
    S_BUF : NETWORK_BUFFER_SHORT;
    R_BUF : NETWORK_BUFFER_SHORT;
    DATA : ARRAY[0..255] OF WORD;
    W_DATA_BITPOS : INT;
    W_DATA_ADR : INT;
    W_POINTS : INT;
    W_ADDR : INT;
    R_DATA_BITPOS : INT;
    R_DATA_ADR : INT;
    R_POINTS : INT;
    R_ADDR : INT;
    FC : INT;
    ENABLE : BOOL;
END_VAR

END_FUNCTION

(* ---- MB_SERVER_DEMO.st ---- *)
FUNCTION MB_SERVER_DEMO
VAR
    IP_CONTROL2_1 : IP_CONTROL2;
    MB_SERVER_1 : MB_SERVER;
    IP_C : IP_C;
    S_BUF : NETWORK_BUFFER_SHORT;
    R_BUF : NETWORK_BUFFER_SHORT;
    DATA : ARRAY[0..255] OF WORD;
    VMAP : ARRAY[1..10] OF VMAP_DATA;
    error : DWORD;
END_VAR

END_FUNCTION

(* ---- MD5_AUX.st ---- *)
FUNCTION MD5_AUX : DWORD
VAR_INPUT
    N : INT;
    A : DWORD;
    B : DWORD;
    C : DWORD;
    D : DWORD;
    X : DWORD;
    U : INT;
    T : DWORD;
END_VAR

VAR
    w : DWORD;
END_VAR
CASE N OF
	1: w := (B AND C) OR (NOT(B) AND D);
	2: w := (B AND D) OR (C AND NOT D);
	3: w := (B XOR C XOR D);
	4: w := (C XOR (B OR  NOT(D)));
END_CASE

MD5_AUX := B + ROL(A + w + X + T,U);

(* revision history

ks	6. dec. 2009 rev 1.0
	original version

*)
END_FUNCTION

(* ---- MD5_CRAM_AUTH_DEMO.st ---- *)
FUNCTION MD5_CRAM_AUTH_DEMO
VAR
    run : BOOL := TRUE;
    timestamp : STRING[64] := 'PDQwMzYuMTA3NjMyNDM4MUBndWlsZGVuc3Rlcm4uemVpdGZvcm0uZGU+';
    password : STRING := 'geheimes_passwort';
    username : STRING := 'benutzer@zeitform.de';
    auth_key : STRING[OSCAT_BASIC.STRING_LENGTH];
    MD5_CRAM_AUTH : MD5_CRAM_AUTH; // Assuming MD5_CRAM_AUTH is a defined derived type
END_VAR

END_FUNCTION

(* ---- MD5_TO_STRH.st ---- *)
FUNCTION MD5_TO_STRH : string
VAR_INPUT
    MD5 : ARRAY[0..15] OF BYTE;
END_VAR

VAR
    i : INT;
    tmp : BYTE;
    pt : POINTER TO BYTE;
END_VAR
pt := ADR(MD5_TO_STRH); (* read output adress to pointer *)

FOR i := 0 TO 15 DO; (* write the 8 hex characters backwards *)
	tmp := SHR(MD5[i],4);
	PT^ := tmp + SEL(tmp <= 9,87,48);
	pt := pt + 1; (* decrement the pointer *)
	tmp := MD5[i] AND 2#1111;
	PT^ := tmp + SEL(tmp <= 9,87,48);
	pt := pt + 1; (* decrement the pointer *)
END_FOR;
pt^:= 0; (* write the closing byte for the string *)

(* revision history

ks	6. dec. 2009 rev 1.0
	original version

*)
END_FUNCTION

(* ---- MID3.st ---- *)
FUNCTION MID3 : REAL
VAR_INPUT
    IN1 : REAL;
    IN2 : REAL;
    IN3 : REAL;
END_VAR
IF IN1 > IN2 THEN MID3 := IN1; IN1 := IN2; IN2 := MID3; END_IF;
IF IN2 > IN3 THEN IN2 := IN3; END_IF;
MID3 := SEL(IN1 > IN2, IN2, IN1);

(*
hm	1.1.2007	rev 1.1
	rewrote the function for better performance

hm	18. mar. 2011	rev 1.2
	improve performance
*)
END_FUNCTION

(* ---- MIN3.st ---- *)
FUNCTION MIN3 : REAL
VAR_INPUT
    in1 : REAL;
    in2 : REAL;
    in3 : REAL;
END_VAR
MIN3 := MIN(MIN(IN1,IN2),IN3);

(* revision history
hm	1.1.2007	rev 1.0
	original release

hm	18. mar. 2011	rev 1.1
	improve performance

*)
END_FUNCTION

(* ---- MINUTE.st ---- *)
FUNCTION MINUTE : INT
VAR_INPUT
    itod : TOD;
END_VAR
MINUTE := DWORD_TO_INT(TOD_TO_DWORD(itod) / 60000 - TOD_TO_DWORD(itod) / 3600000 * 60);

(* change history

2.10.2006 changes name of input to itod

*)
END_FUNCTION

(* ---- MINUTE_OF_DT.st ---- *)
FUNCTION MINUTE_OF_DT : INT
VAR_INPUT
    XDT : DT;
END_VAR
MINUTE_OF_DT := DWORD_TO_INT(DT_TO_DWORD(XDT) MOD 3600) / 60;

(* revision history
hm		6.9.2008	rev 1.0
	original version

*)
END_FUNCTION

(* ---- MINUTE_TO_TIME.st ---- *)
FUNCTION MINUTE_TO_TIME : TIME
VAR_INPUT
    IN : REAL;
END_VAR
MINUTE_TO_TIME := DWORD_TO_TIME(REAL_TO_DWORD(IN * 60000.0));

(* revision history
hm	4. aug 2006	rev 1.0
	original version

hm	14. mar 2008	rev 1.1
	rounded the input after the last digit

hm	24. feb. 2009	rev 1.2
	changed input to IN

*)
END_FUNCTION

(* ---- MIRROR.st ---- *)
FUNCTION MIRROR : string
VAR_INPUT
    str: STRING(STRING_LENGTH);
END_VAR

VAR
    pi: POINTER TO ARRAY[1..255] OF BYTE;
    po: POINTER TO BYTE;
    lx: INT;
    i: INT;
END_VAR
pi := ADR(str);
po := ADR(mirror);
lx := LEN(str);
FOR i := lx TO 1 BY - 1 DO
	po^ := pi^[i];
	po := po + 1;
END_FOR;
(* close output string *)
po^:= 0;

(* revision histroy
hm	4. feb. 2008	rev 1.0
	original release

hm	29. mar. 2008	rev 1.1
	changed STRING to STRING(STRING_LENGTH)
*)
END_FUNCTION

(* ---- MIX.st ---- *)
FUNCTION MIX : REAL
VAR_INPUT
    A : REAL;
    B : REAL;
    M : REAL;
END_VAR
MIX := (1.0 - M) * A + M * B;

(* revision history
hm	19. Nov 2007	rev 1.0
	original version

hm	10. mar 2009	rev 1.1
	real constants updated to new systax using dot

*)
END_FUNCTION

(* ---- MODR.st ---- *)
FUNCTION MODR : REAL
VAR_INPUT
    IN : REAL;
    DIVI : REAL;
END_VAR
IF divi = 0.0 THEN
	MODR := 0.0;
ELSE
	MODR := in - DINT_TO_REAL(FLOOR2(in / divi)) * divi;
END_IF;

(* revision history

hm	4. aug.2006		rev 1.0

hm	28. jan.2007	rev 1.1
	modr(x,0) will deliver the result 0

hm	21. mar 2008	rev 1.2
	use D_trunc for compatibility reasons

hm	4. apr. 2008	rev 1.3
	added type conversion to avoid warnings under codesys 3.0

hm	31. oct. 2008	rev 1.4
	changed algorithm to the more common version using floor instead of TRUNC

hm	10. mar. 2009	rev 1.5
	real constants updated to new systax using dot

*)
END_FUNCTION

(* ---- MONTH_BEGIN.st ---- *)
FUNCTION MONTH_BEGIN : DATE
VAR_INPUT
    idate : DATE;
END_VAR
MONTH_BEGIN := DWORD_TO_DATE(DATE_TO_DWORD(idate) - INT_TO_DWORD(DAY_OF_MONTH(idate) - 1) * 86400);

(* revision history
hm	15. jun. 2008	rev 1.0
	original version

*)
END_FUNCTION

(* ---- MONTH_END.st ---- *)
FUNCTION MONTH_END : DATE
VAR_INPUT
    IDATE : DATE;
END_VAR
MONTH_END := DWORD_TO_DATE(DATE_TO_DWORD(SET_DATE(YEAR_OF_DATE(idate),MONTH_OF_DATE(idate)+1,1)) - 86400);

(* revision history
hm	15. jun. 2008	rev 1.0
	original version

hm	7. oct. 2008	rev 1.1
	changed function year to year_of_date
	changed function month to month_of_date

*)
END_FUNCTION

(* ---- MONTH_OF_DATE.st ---- *)
FUNCTION MONTH_OF_DATE : INT
VAR_INPUT
    IDATE: DATE;
END_VAR
MONTH_OF_DATE := DAY_OF_YEAR(idate);
IF MONTH_OF_DATE < 32 THEN
	MONTH_OF_DATE := 1;
ELSIF LEAP_OF_DATE(IDATE) THEN
	MONTH_OF_DATE := (MONTH_OF_DATE * 53 + 1668) / 1623;
ELSE
	MONTH_OF_DATE := (MONTH_OF_DATE * 53 + 1700) / 1620;
END_IF;

(* code for rev 1.2
MONTH_OF_DATE := DAY_OF_YEAR(IDATE);
IF LEAP_OF_DATE(IDATE) THEN
	CASE MONTH_OF_DATE OF
		1..31 	:	MONTH_OF_DATE := 1;
		32..60	:	MONTH_OF_DATE := 2;
		61..91	:	MONTH_OF_DATE := 3;
		92..121 :	MONTH_OF_DATE := 4;
		122..152:	MONTH_OF_DATE := 5;
		153..182:	MONTH_OF_DATE := 6;
		183..213:	MONTH_OF_DATE := 7;
		214..244:	MONTH_OF_DATE := 8;
		245..274:	MONTH_OF_DATE := 9;
		275..305:	MONTH_OF_DATE := 10;
		306..335:	MONTH_OF_DATE := 11;
		336..366:	MONTH_OF_DATE := 12;
	END_CASE;
ELSE
	CASE MONTH_OF_DATE OF
		1..31 	:	MONTH_OF_DATE := 1;
		32..59	:	MONTH_OF_DATE := 2;
		60..90	:	MONTH_OF_DATE := 3;
		91..120 :	MONTH_OF_DATE := 4;
		121..151:	MONTH_OF_DATE := 5;
		152..181:	MONTH_OF_DATE := 6;
		182..212:	MONTH_OF_DATE := 7;
		213..243:	MONTH_OF_DATE := 8;
		244..273:	MONTH_OF_DATE := 9;
		274..304:	MONTH_OF_DATE := 10;
		305..334:	MONTH_OF_DATE := 11;
		335..365:	MONTH_OF_DATE := 12;
	END_CASE;
END_IF;
*)

(* revision history
hm	1. aug 2006	rev 1.0
	original version

hm	1. okt 2007	rev 1.1
	replaced old code (string conversion) with mathematics
	the execution time is now multiple times faster.

hm	7. oct. 2008	rev 1.2
	changed name of function from month to MONTH_OF_DATE

hm	27. mar. 2009	rev 1.3
	new improved code

*)
END_FUNCTION

(* ---- MONTH_TO_STRING.st ---- *)
FUNCTION MONTH_TO_STRING : string
VAR_INPUT
    MTH : INT;
    LANG : INT;
    LX : INT;
END_VAR

VAR
    ly : INT;
END_VAR
IF LANG <= 0 THEN Ly := LANGUAGE.DEFAULT; ELSE ly := MIN(LANG, language.LMAX); END_IF;
IF MTH < 1 OR MTH > 12 THEN
	RETURN;
ELSIF LX = 0 THEN
	MONTH_TO_STRING := language.MONTHS[ly, MTH];
ELSIF Lx = 3 THEN
	MONTH_TO_STRING := language.MONTHS3[ly, MTH];
END_IF;

(* revisison history

hm	21. sep. 2008	rev 1.0
	original version

hm	19. oct. 2008	rev 1.1
	changed language setup constants

hm 16.  jul 2024   rev 1.2
       addaed boundary check to respect array limits
*)
END_FUNCTION

(* ---- MS_TO_BFT.st ---- *)
FUNCTION MS_TO_BFT : INT
VAR_INPUT
    MS : REAL;
END_VAR
MS_TO_BFT := REAL_TO_INT(EXPT(MS * 1.196172, 0.666667));

(* revision history
hm	12. 6. 2008		rev 1.0
	original version

*)
END_FUNCTION

(* ---- MS_TO_KMH.st ---- *)
FUNCTION MS_TO_KMH : REAL
VAR_INPUT
    ms : REAL;
END_VAR
MS_TO_KMH := ms * 3.6;
END_FUNCTION

(* ---- MUL_ADD.st ---- *)
FUNCTION MUL_ADD : REAL
VAR_INPUT
    X : REAL;
    K : REAL;
    O : REAL;
END_VAR
MUL_ADD := X * K + O;

(* revision history
hm	28. feb 2007
	original version

hm	11.nov 2007		rev 1.1
	deleted preset values for K and O this makes no sense for a function

*)
END_FUNCTION

(* ---- MULTI_IN.st ---- *)
FUNCTION MULTI_IN : REAL
VAR_INPUT
    in_1 : REAL;
    in_2 : REAL;
    in_3 : REAL;
    default : REAL;
    in_min : REAL;
    in_max : REAL;
    mode : BYTE;
END_VAR

VAR
    count : INT;
    F1 : BOOL;
    F2 : BOOL;
    F3 : BOOL;
END_VAR
F1 :=  in_1 > in_min AND in_1 < in_max;
F2 :=  in_2 > in_min AND in_2 < in_max;
F3 :=  in_3 > in_min AND in_3 < in_max;

CASE mode OF
0:	count := 0;
	IF F1 THEN
		count := count + 1;
		MULTI_IN := in_1;
	ELSE
		MULTI_IN := 0.0;
	END_IF;
	IF F2 THEN
		count := count + 1;
		MULTI_IN := MULTI_IN + in_2;
	END_IF;
	IF F3 THEN
		count := count + 1;
		MULTI_IN := MULTI_IN + in_3;
	END_IF;
	MULTI_IN := SEL(count = 0, MULTI_IN / INT_TO_REAL(count), default);

1:	MULTI_IN := SEL(F1, default, IN_1);

2:	MULTI_IN := SEL(F2, default, IN_2);

3:	MULTI_IN := SEL(F3, default, IN_3);

4:	MULTI_IN := default;

5:	MULTI_IN := SEL(F1, in_max, IN_1);
	IF F2 AND in_2 < MULTI_IN THEN MULTI_IN := in_2; END_IF;
	IF F3 AND in_3 < MULTI_IN THEN MULTI_IN := in_3; END_IF;
	IF MULTI_IN = in_max THEN MULTI_IN := default; END_IF;

6:	MULTI_IN := SEL(F1, in_min, IN_1);
	IF F2 AND in_2 > MULTI_IN THEN MULTI_IN := in_2; END_IF;
	IF F3 AND in_3 > MULTI_IN THEN MULTI_IN := in_3; END_IF;
	IF MULTI_IN = in_min THEN MULTI_IN := default; END_IF;

7:	IF F1 AND F2 AND F3 THEN MULTI_IN := MID3(in_1, in_2, in_3);
	ELSIF F1 AND F2 THEN MULTI_IN := MIN(in_1, in_2);
	ELSIF F1 AND F3 THEN MULTI_IN := MIN(in_1, in_3);
	ELSIF F2 AND F3 THEN MULTI_IN := MIN(in_2, in_3);
	ELSIF F1 THEN MULTI_IN := in_1;
	ELSIF F2 THEN MULTI_IN := in_2;
	ELSIF F3 THEN MULTI_IN := in_3;
	ELSE MULTI_IN := default;
	END_IF;

END_CASE;

(*
hm 1.1.2007		rev 1.1
	changed midr to mid3 function

hm	14. 10. 2008	rev 1.2
	corrected an error for in_3 overrange detection
	improved performance

hm	11. mar. 2009	rev 1.3
	changed real constants to use dot syntax

hm	18. jul. 2009	rev 1.4
	improved performance
*)
END_FUNCTION

(* ---- MULTIME.st ---- *)
FUNCTION MULTIME : TIME
VAR_INPUT
    t : TIME;
    M : REAL;
END_VAR
MULTIME := DWORD_TO_TIME(REAL_TO_DWORD(DWORD_TO_REAL(TIME_TO_DWORD(t))*M));

(* revision history
hm		2. oct 2006	rev 1.0
	original version

hm		14. mar 2008	rev 1.1
	rounded the result after the last digit

*)
END_FUNCTION

(* ---- MUX_2.st ---- *)
FUNCTION MUX_2 : BOOL
VAR_INPUT
    D0 : BOOL;
    D1 : BOOL;
    A0 : BOOL;
END_VAR
MUX_2 := SEL(A0, D0, D1);

(*
revision history:
hm	5.10.2006		rev 1.1
	changed to ST Langage for better portability.

hm	16. oct. 2008	rev 1.2
	improved performance

*)
END_FUNCTION

(* ---- MUX_4.st ---- *)
FUNCTION MUX_4 : BOOL
VAR_INPUT
    D0 : BOOL;
    D1 : BOOL;
    D2 : BOOL;
    D3 : BOOL;
    A0 : BOOL;
    A1 : BOOL;
END_VAR
IF A1 THEN
	MUX_4 := SEL(A0, D2, D3);
ELSE
	MUX_4 := SEL(A0, D0, D1);
END_IF;

(*
revision history:
hm 	5.10.2006		rev 1.1
	rewritten to ST for better portability

hm	16. oct. 2008	rev 1.2
	improved performance

*)
END_FUNCTION

(* ---- MUX_R2.st ---- *)
FUNCTION MUX_R2 : REAL
VAR_INPUT
    IN0 : REAL;
    IN1 : REAL;
    A : BOOL;
END_VAR
MUX_R2 := SEL(A, IN0, IN1);

(* revision history
hm	19. jan. 2007	rev 1.0
	original version

hm	16. oct. 2008	rev 1.1
	improved performance

*)
END_FUNCTION

(* ---- MUX_R4.st ---- *)
FUNCTION MUX_R4 : REAL
VAR_INPUT
    IN0 : REAL;
    IN1 : REAL;
    IN2 : REAL;
    IN3 : REAL;
    A0 : BOOL;
    A1 : BOOL;
END_VAR
IF A1 THEN
	MUX_R4 := SEL(A0, IN2, IN3);
ELSE
	MUX_R4 := SEL(A0, IN0, IN1);
END_IF;

(* revision history
hm	19. jan 2007	rev 1.0
	original version

hm	16. oct. 2008	rev 1.1
	improved performance
*)
END_FUNCTION

(* ---- NEGX.st ---- *)
FUNCTION NEGX : REAL
VAR_INPUT
    X : REAL;
END_VAR
NEGX := -X;

(* revision history
hm	26. oct. 2008	rev 1.0
	original version

*)
END_FUNCTION

(* ---- NET_VAR_MASTER_DEMO.st ---- *)
FUNCTION NET_VAR_MASTER_DEMO
VAR
    NET_VAR_CONTROL_1 : NET_VAR_CONTROL;
    activate : BOOL := TRUE;
    run : BOOL;
    udp : BOOL := TRUE;
    master : BOOL := TRUE;
    remote_port : WORD := 10000;
    scan_time : TIME := TIME#1s0ms;
    watchdog : TIME := TIME#2s0ms;
    error : DWORD;
    x : NET_VAR_DATA;
    NET_VAR_BOOL8_1 : NET_VAR_BOOL8;
    id_b8 : BYTE;
    in_b1 : BOOL;
    in_b2 : BOOL;
    in_b3 : BOOL;
    in_b4 : BOOL;
    in_b5 : BOOL;
    in_b6 : BOOL;
    in_b7 : BOOL;
    in_b8 : BOOL;
    out_b1 : BOOL;
    out_b2 : BOOL;
    out_b3 : BOOL;
    out_b4 : BOOL;
    out_b5 : BOOL;
    out_b6 : BOOL;
    out_b7 : BOOL;
    out_b8 : BOOL;
    NET_VAR_STRING_1 : NET_VAR_STRING;
    in_s1 : STRING( OSCT_BASIC.STRING_LENGTH );
    out_s1 : STRING( OSCT_BASIC.STRING_LENGTH );
    id_s : BYTE;
    NET_VAR_BUFFER_1 : NET_VAR_BUFFER;
    id_bu : BYTE;
    BUF_IN : ARRAY[1..64] OF BYTE;
    BUF_OUT : ARRAY[1..64] OF BYTE;
    id_dw : BYTE;
    NET_VAR_DWORD8_1 : NET_VAR_DWORD8;
    in_dw1 : DWORD;
    in_dw2 : DWORD;
    in_dw3 : DWORD;
    in_dw4 : DWORD;
    in_dw5 : DWORD;
    in_dw6 : DWORD;
    in_dw7 : DWORD;
    in_dw8 : DWORD;
    out_dw1 : DWORD;
    out_dw2 : DWORD;
    out_dw3 : DWORD;
    out_dw4 : DWORD;
    out_dw5 : DWORD;
    out_dw6 : DWORD;
    out_dw7 : DWORD;
    out_dw8 : DWORD;
    NET_VAR_REAL8_1 : NET_VAR_REAL8;
    in_r1 : REAL;
    in_r2 : REAL;
    in_r3 : REAL;
    in_r4 : REAL;
    in_r5 : REAL;
    in_r6 : REAL;
    in_r7 : REAL;
    in_r8 : REAL;
    out_r1 : REAL;
    out_r2 : REAL;
    out_r3 : REAL;
    out_r4 : REAL;
    out_r5 : REAL;
    out_r6 : REAL;
    out_r7 : REAL;
    out_r8 : REAL;
    id_r : BYTE;
    NET_VAR_X8_1 : NET_VAR_X8;
    in_x_re1 : REAL;
    in_x_re2 : REAL;
    in_x_di1 : DINT;
    in_x_di2 : DINT;
    in_x_ud1 : UDINT;
    in_x_ud2 : UDINT;
    in_x_dw1 : DWORD;
    in_x_dw2 : DWORD;
    out_x_re1 : REAL;
    out_x_re2 : REAL;
    out_x_di1 : DINT;
    out_x_di2 : DINT;
    out_x_ud1 : UDINT;
    out_x_ud2 : UDINT;
    out_x_dw1 : DWORD;
    out_x_dw2 : DWORD;
    id_x8 : BYTE;
END_VAR

END_FUNCTION

(* ---- NET_VAR_SLAVE_DEMO.st ---- *)
FUNCTION NET_VAR_SLAVE_DEMO
VAR
    NET_VAR_CONTROL_1 : NET_VAR_CONTROL;
    activate : BOOL := TRUE;
    run : BOOL;
    udp : BOOL := TRUE;
    master : BOOL := FALSE;
    remote_port : WORD := 10000;
    scan_time : TIME := TIME#1s0ms;
    watchdog : TIME := TIME#2s0ms;
    error : DWORD;
    x : NET_VAR_DATA;
    NET_VAR_BOOL8_1 : NET_VAR_BOOL8;
    id_b8 : BYTE;
    in_b1 : BOOL;
    in_b2 : BOOL;
    in_b3 : BOOL;
    in_b4 : BOOL;
    in_b5 : BOOL;
    in_b6 : BOOL;
    in_b7 : BOOL;
    in_b8 : BOOL;
    out_b1 : BOOL;
    out_b2 : BOOL;
    out_b3 : BOOL;
    out_b4 : BOOL;
    out_b5 : BOOL;
    out_b6 : BOOL;
    out_b7 : BOOL;
    out_b8 : BOOL;
    NET_VAR_STRING_1 : NET_VAR_STRING;
    in_s1 : STRING[OSCAT_BASIC.STRING_LENGTH];
    out_s1 : STRING[OSCAT_BASIC.STRING_LENGTH];
    id_s : BYTE;
    NET_VAR_BUFFER_1 : NET_VAR_BUFFER;
    id_bu : BYTE;
    BUF_IN : ARRAY[1..64] OF BYTE;
    BUF_OUT : ARRAY[1..64] OF BYTE;
    id_dw : BYTE;
    NET_VAR_DWORD8_1 : NET_VAR_DWORD8;
    in_dw1 : DWORD;
    in_dw2 : DWORD;
    in_dw3 : DWORD;
    in_dw4 : DWORD;
    in_dw5 : DWORD;
    in_dw6 : DWORD;
    in_dw7 : DWORD;
    in_dw8 : DWORD;
    out_dw1 : DWORD;
    out_dw2 : DWORD;
    out_dw3 : DWORD;
    out_dw4 : DWORD;
    out_dw5 : DWORD;
    out_dw6 : DWORD;
    out_dw7 : DWORD;
    out_dw8 : DWORD;
    NET_VAR_REAL8_1 : NET_VAR_REAL8;
    in_r1 : REAL;
    in_r2 : REAL;
    in_r3 : REAL;
    in_r4 : REAL;
    in_r5 : REAL;
    in_r6 : REAL;
    in_r7 : REAL;
    in_r8 : REAL;
    out_r1 : REAL;
    out_r2 : REAL;
    out_r3 : REAL;
    out_r4 : REAL;
    out_r5 : REAL;
    out_r6 : REAL;
    out_r7 : REAL;
    out_r8 : REAL;
    id_r : BYTE;
    NET_VAR_X8_1 : NET_VAR_X8;
    in_x_re1 : REAL;
    in_x_re2 : REAL;
    in_x_di1 : DINT;
    in_x_di2 : DINT;
    in_x_ud1 : UDINT;
    in_x_ud2 : UDINT;
    in_x_dw1 : DWORD;
    in_x_dw2 : DWORD;
    out_x_re1 : REAL;
    out_x_re2 : REAL;
    out_x_di1 : DINT;
    out_x_di2 : DINT;
    out_x_ud1 : UDINT;
    out_x_ud2 : UDINT;
    out_x_dw1 : DWORD;
    out_x_dw2 : DWORD;
    id_x8 : BYTE;
END_VAR

END_FUNCTION

(* ---- NETWORK_VERSION.st ---- *)
FUNCTION NETWORK_VERSION : DWORD
VAR_INPUT
    IN : BOOL;
END_VAR
IF in THEN
	NETWORK_VERSION := DATE_TO_DWORD(D#2016-07-01);
ELSE
	NETWORK_VERSION := 135;
END_IF;

(* revision history
ks	2. feb 2011	rev 1.0
	original version

*)
END_FUNCTION

(* ---- OCT_TO_BYTE.st ---- *)
FUNCTION OCT_TO_BYTE : BYTE
VAR_INPUT
    OCT : STRING[10];
END_VAR

VAR
    pt : POINTER TO BYTE;
    i : INT;
    X : BYTE;
    stop : INT;
END_VAR
pt := ADR(oct);
stop := LEN(oct);
FOR I := 1 TO stop DO
	(* read the first character and subtract 48 to get value in decimal 0 = 48 *)
	x := pt^;
	(* calculate the value of the digit *)
	IF X > 47 AND x < 56 THEN
		OCT_TO_BYTE := SHL(OCT_TO_BYTE,3) + X - 48;
	END_IF;
	pt := pt + 1;
END_FOR;

(* revision histroy
hm	18. jun. 2008	rev 1.0
	original release

hm	20. sep. 2008	rev 1.1
	changed length of input string from 20 to 10

*)
END_FUNCTION

(* ---- OCT_TO_DWORD.st ---- *)
FUNCTION OCT_TO_DWORD : DWORD
VAR_INPUT
    OCT : STRING[20];
END_VAR

VAR
    pt : POINTER TO BYTE;
    i : INT;
    X : BYTE;
    stop : INT;
END_VAR
pt := ADR(oct);
stop := LEN(oct);
FOR I := 1 TO stop DO
	(* read the first character and subtract 48 to get value in decimal 0 = 48 *)
	x := pt^;
	(* calculate the value of the digit *)
	IF X > 47 AND x < 56 THEN
		OCT_TO_DWORD := SHL(OCT_TO_DWORD,3) + X - 48;
	END_IF;
	pt := pt + 1;
END_FOR;

(* revision histroy
hm	18. jun. 2008	rev 1.0
	original release

*)
END_FUNCTION

(* ---- OFFSET.st ---- *)
FUNCTION OFFSET : REAL
VAR_INPUT
    X : REAL;
    O1 : BOOL;
    O2 : BOOL;
    O3 : BOOL;
    O4 : BOOL;
    D : BOOL;
    Offset_1 : REAL;
    Offset_2 : REAL;
    Offset_3 : REAL;
    Offset_4 : REAL;
    default : REAL;
END_VAR
IF D THEN OFFSET := default; ELSE OFFSET := X; END_IF;
IF O1 THEN OFFSET := OFFSET + offset_1; END_IF;
IF O2 THEN OFFSET := OFFSET + offset_2; END_IF;
IF O3 THEN OFFSET := OFFSET + offset_3; END_IF;
IF O4 THEN OFFSET := OFFSET + offset_4; END_IF;

(* revision history
hm	12. jan 2007
	original version

*)
END_FUNCTION

(* ---- OFFSET2.st ---- *)
FUNCTION OFFSET2 : REAL
VAR_INPUT
    X : REAL;
    O1 : BOOL;
    O2 : BOOL;
    O3 : BOOL;
    O4 : BOOL;
    D : BOOL;
    Offset_1 : REAL;
    Offset_2 : REAL;
    Offset_3 : REAL;
    Offset_4 : REAL;
    default : REAL;
END_VAR
IF D THEN OFFSET2 := default; ELSE OFFSET2 := X; END_IF;
IF O4 THEN OFFSET2 := OFFSET2 + offset_4;
ELSIF O3 THEN OFFSET2 := OFFSET2 + offset_3;
ELSIF O2 THEN OFFSET2 := OFFSET2 + offset_2;
ELSIF O1 THEN OFFSET2 := OFFSET2 + offset_1;
END_IF;
END_FUNCTION

(* ---- OM_TO_F.st ---- *)
FUNCTION OM_TO_F : REAL
VAR_INPUT
    OM : REAL;
END_VAR
OM_TO_F := OM / math.PI2;

(* revision history
hm	22. jan. 2007	rev 1.0
	original version

hm	18. oct. 2008	rev 1.1
	using math constants

*)
END_FUNCTION

(* ---- OSCAT_VERSION.st ---- *)
FUNCTION OSCAT_VERSION : DWORD
VAR_INPUT
    IN : BOOL;
END_VAR
IF in THEN
	OSCAT_VERSION := DATE_TO_DWORD(D#2024-07-16);
ELSE
	OSCAT_VERSION := 335;
END_IF;

(* revision history
hm	6. oct 2006	rev 1.0
	original version

hm	16. dec 2007	rev 1.1
	added possibility to return date and version depending on IN.

*)
END_FUNCTION

(* ---- OVERRIDE.st ---- *)
FUNCTION OVERRIDE : REAL
VAR_INPUT
    X1 : REAL;
    X2 : REAL;
    X3 : REAL;
    E1 : BOOL;
    E2 : BOOL;
    E3 : BOOL;
END_VAR
IF E1 THEN OVERRIDE := X1; END_IF;
IF E2 AND ABS(x2) > ABS(OVERRIDE) THEN OVERRIDE := X2; END_IF;
IF E3 AND ABS(x3) > ABS(OVERRIDE) THEN OVERRIDE := X3; END_IF;

(* revision history
hm	4.11.2007		rev 1.0
	original version

*)
END_FUNCTION

(* ---- PARITY.st ---- *)
FUNCTION PARITY : BOOL
VAR_INPUT
    in : DWORD;
END_VAR
WHILE in > 0 DO
	PARITY := PARITY XOR in.0 XOR in.1 XOR in.2 XOR in.3;
	in := SHR(in,4);
END_WHILE;

(* code before rev 1.2
WHILE in > 0 DO
	IF in.0 THEN cnt := cnt +1; END_IF;
	in := SHR(in,1);
END_WHILE;
IF (cnt MOD 2) = 1 THEN parity := TRUE; ELSE parity := FALSE; END_IF;
*)

(* revision history

rev 1.0 hm 1 sep 2006
	original version

rev 1.1 hm 10.9.2007
	changed algorithm to improve performance

rev 1.2	hm	8 dec 2007
	changed algorithm to improve performance

rev 1.3	hm	18 feb 2008
	changed algorithm to improve performance
*)
END_FUNCTION

(* ---- PERIOD.st ---- *)
FUNCTION PERIOD : BOOL
VAR_INPUT
    d1: DATE;
    dx: DATE;
    d2: DATE;
END_VAR

VAR
    day1: INT;
    day2: INT;
    dayx: INT;
END_VAR
day1 := DAY_OF_YEAR(d1);
day2 := DAY_OF_YEAR(d2);
dayx := DAY_OF_YEAR(dx);
IF NOT LEAP_OF_DATE(dx) AND dayx > 58 THEN dayx := dayx + 1; END_IF;
IF NOT LEAP_OF_DATE(d1) AND day1 > 58 THEN day1 := day1 + 1; END_IF;
IF NOT LEAP_OF_DATE(d2) AND day2 > 58 THEN day2 := day2 + 1; END_IF;

IF day2 < day1 THEN
	(* the period spans over the new year *)
	PERIOD := dayx <= day2 OR dayx >= day1;
ELSE
	PERIOD := dayx >= day1 AND dayx <= day2;
END_IF;

(* code before rev 1.2
yx := year(dx);
p1 := date_add(d1,0,0,0,yx - year(d1));
p2 := date_add(d2,0,0,0,yx - year(d2));

IF p2 >= p1 THEN
	period := dx <= p2  AND dx >= p1;
ELSE
	period := dx <= p2 OR dx >= p1;
END_IF;
*)

(* revision history

hm		19. sep 2007	rev 1.0
	original version

hm		20. sep 2007	rev 1.1
	corrected a problem with leap year

hm		4. jan 2008		rev 1.2
	changed code for better performance

hm		22. mar. 2008	rev 1.3
	function would deliver wrong results when d1, d2 or dx are a leap_year

*)
END_FUNCTION

(* ---- PERIOD2.st ---- *)
FUNCTION PERIOD2 : BOOL
VAR_INPUT
    DP : ARRAY[0..3, 0..1] OF DATE; // Array of DATEs
    DX : DATE;                     // Single DATE
END_VAR
PERIOD2 := 	(DX >= DP[0,0] AND DX <= DP[0,1]) OR
			(DX >= DP[1,0] AND DX <= DP[1,1]) OR
			(DX >= DP[2,0] AND DX <= DP[2,1]) OR
			(DX >= DP[3,0] AND DX <= DP[3,1]);

(* revision history

hm		27. apr 2008	rev 1.0
	original version

*)
END_FUNCTION
